   // ---------- 网络 3 ----------
   // 标题：******************************         Total Cmd . Start      ********************************
   // 含义：将 ((#Cmd.Man.StartTest OR #Step.Main.Start) AND #ManMode) AND NOT (#Step.Main.End) 赋给 #Step.Main.Start
   #Step.Main.Start := ((#Cmd.Man.StartTest OR #Step.Main.Start) AND #ManMode) AND NOT (#Step.Main.End);
   // 含义：将 ((#Cmd.Man.StartTest OR #Step.Main.Start) AND #ManMode) AND NOT (#Step.Main.End) 赋给 #Status.Busy
   #Status.Busy := ((#Cmd.Man.StartTest OR #Step.Main.Start) AND #ManMode) AND NOT (#Step.Main.End);
   // 含义：条件 NOT (((#Cmd.Man.StartTest OR #Step.Main.Start) AND #ManMode) AND NOT (#Step.Main.End)) 成立时，将 FALSE 传送到 #Status.TaskDone
   IF NOT (((#Cmd.Man.StartTest OR #Step.Main.Start) AND #ManMode) AND NOT (#Step.Main.End)) THEN
       #Status.TaskDone := FALSE;
   END_IF;
   // 含义：条件 NOT (((#Cmd.Man.StartTest OR #Step.Main.Start) AND #ManMode) AND NOT (#Step.Main.End)) 成立时，将 FALSE 传送到 #Step.Main.ErrEnd
   IF NOT (((#Cmd.Man.StartTest OR #Step.Main.Start) AND #ManMode) AND NOT (#Step.Main.End)) THEN
       #Step.Main.ErrEnd := FALSE;
   END_IF;
   // 含义：条件 NOT (((#Cmd.Man.StartTest OR #Step.Main.Start) AND #ManMode) AND NOT (#Step.Main.End)) 成立时，将 0 传送到 #Step.RandomStepNO
   IF NOT (((#Cmd.Man.StartTest OR #Step.Main.Start) AND #ManMode) AND NOT (#Step.Main.End)) THEN
       #Step.RandomStepNO := 0;
   END_IF;

   // ---------- 网络 4 ----------
   // 标题：TimeOut
   // 含义：条件 #Status.Busy AND NOT (#Step.Main.S1) 成立时，将 FALSE 传送到 #Timer_TimeOut.IN
   IF #Status.Busy AND NOT (#Step.Main.S1) THEN
       #Timer_TimeOut.IN := FALSE;
   END_IF;
   // 含义：调用定时器实例 #Timer_TimeOut
   #Timer_TimeOut(TV := #Ctrl_IN.InitParameter.TimeOutSetValue);
   // 含义：当 #Status.Busy 为 TRUE 时置位 #Timer_TimeOut.IN，否则复位（触点→线圈）
   IF #Status.Busy THEN
       #Timer_TimeOut.IN := TRUE;
   ELSE
       #Timer_TimeOut.IN := FALSE;
   END_IF;
   // 含义：条件 #Status.Busy AND #Step.Main.RandomTestCycleReStart 成立时，将 "SyS_Time" 传送到 #Aux.CycleTime_StartTime
   IF #Status.Busy AND #Step.Main.RandomTestCycleReStart THEN
       #Aux.CycleTime_StartTime := "SyS_Time";
   END_IF;
   // 含义：条件 #Status.Busy 成立时，将 ("SyS_Time" - #Aux.CycleTime_StartTime) 传送到 #Ctrl_Out.LastCylceTime
   IF #Status.Busy THEN
       #Ctrl_Out.LastCylceTime := ("SyS_Time" - #Aux.CycleTime_StartTime);
   END_IF;

   // ---------- 网络 5 ----------
   // 标题：Init
   // 含义：条件 #Step.Main.Start AND NOT (#Step.Main.S1) 成立时，将 TRUE 传送到 #Step.Main.RandomTestCycleReStart
   IF #Step.Main.Start AND NOT (#Step.Main.S1) THEN
       #Step.Main.RandomTestCycleReStart := TRUE;
   END_IF;
   // 含义：条件 #Step.Main.Start AND NOT (#Step.Main.S1) 成立时，将 #Servo_CTRL_IN.InitParameter.TimeOutSetValue 传送到 #Aux.TimeOutSetValue
   IF #Step.Main.Start AND NOT (#Step.Main.S1) THEN
       #Aux.TimeOutSetValue := #Servo_CTRL_IN.InitParameter.TimeOutSetValue;
   END_IF;
   // 含义：条件 #Step.Main.Start AND NOT (#Step.Main.S1) 成立时，将 t#15d 传送到 #Servo_CTRL_IN.InitParameter.TimeOutSetValue
   IF #Step.Main.Start AND NOT (#Step.Main.S1) THEN
       #Servo_CTRL_IN.InitParameter.TimeOutSetValue := t#15d;
   END_IF;
   // 含义：条件 #Step.Main.Start AND NOT (#Step.Main.S1) 成立时，将 0 传送到 #Ctrl_Out.AcutalCycleCounter
   IF #Step.Main.Start AND NOT (#Step.Main.S1) THEN
       #Ctrl_Out.AcutalCycleCounter := 0;
   END_IF;
   // 含义：条件 #Step.Main.Start AND NOT (#Step.Main.S1) 成立时，将 0 传送到 #Step.RandomStepNO
   IF #Step.Main.Start AND NOT (#Step.Main.S1) THEN
       #Step.RandomStepNO := 0;
   END_IF;
   // 含义：当 #Step.Main.Start 为 TRUE 时置位 #Step.Main.S1，否则复位（触点→线圈）
   IF #Step.Main.Start THEN
       #Step.Main.S1 := TRUE;
   ELSE
       #Step.Main.S1 := FALSE;
   END_IF;

   // ---------- 网络 6 ----------
   // 标题：***************************以上无需修改  ********************************
   // （空白网络）

   // ---------- 网络 7 ----------
   // 标题：乱序随机测试---随机数的生成；
   // 含义：条件 #Step.Main.RandomTestCycleReStart 成立时，将 #Step.RandomStepNO 传送到 #Ctrl_Out.LastStep
   IF #Step.Main.RandomTestCycleReStart THEN
       #Ctrl_Out.LastStep := #Step.RandomStepNO;
   END_IF;
   // 含义：条件 #Step.Main.RandomTestCycleReStart 成立时，将 (TOD_TO_DINT("SyS_Time") MOD 2) 传送到 #T_DINT
   IF #Step.Main.RandomTestCycleReStart THEN
       #T_DINT := (TOD_TO_DINT("SyS_Time") MOD 2);
   END_IF;
   // 含义：条件 #Step.Main.RandomTestCycleReStart 成立时，将 #T_DINT 传送到 #Step.RandomStepNO
   IF #Step.Main.RandomTestCycleReStart THEN
       #Step.RandomStepNO := #T_DINT;
   END_IF;
   // 含义：条件 #Step.Main.RandomTestCycleReStart 成立时，将 FALSE 传送到 #Status.TaskDone
   IF #Step.Main.RandomTestCycleReStart THEN
       #Status.TaskDone := FALSE;
   END_IF;
   // 含义：条件 #Step.Main.RandomTestCycleReStart 成立时，将 FALSE 传送到 #Status.TaskIO
   IF #Step.Main.RandomTestCycleReStart THEN
       #Status.TaskIO := FALSE;
   END_IF;

   // ---------- 网络 8 ----------
   // 标题：根据随机数进行跳转；
   // JmpList resolved

   // ---------- 网络 9 ----------
   // 标题：#Step.RandomStepNO  = 0:
   // 含义：将 ((((#Step.Main.Start AND (#Step.RandomStepNO = 0))) AND NOT (#Step.Main.RandomTestCycleReStart)) AND NOT (#Servo_Status.Busy)) OR ((((#Step.Main.Start AND (#Step.RandomStepNO = 0))) AND NOT (#Step.Main.RandomTestCycleReStart)) AND #Step.Main.S10) 赋给 #Step.Main.S10
   #Step.Main.S10 := ((((#Step.Main.Start AND (#Step.RandomStepNO = 0))) AND NOT (#Step.Main.RandomTestCycleReStart)) AND NOT (#Servo_Status.Busy)) OR ((((#Step.Main.Start AND (#Step.RandomStepNO = 0))) AND NOT (#Step.Main.RandomTestCycleReStart)) AND #Step.Main.S10);
   // 含义：条件 ((((#Step.Main.Start AND (#Step.RandomStepNO = 0))) AND NOT (#Step.Main.RandomTestCycleReStart)) AND #Step.Main.S10) AND NOT (#Step.Main.S11) 成立时，将 TRUE 传送到 #Servo_Cmd.Auto.StartTask
   IF ((((#Step.Main.Start AND (#Step.RandomStepNO = 0))) AND NOT (#Step.Main.RandomTestCycleReStart)) AND #Step.Main.S10) AND NOT (#Step.Main.S11) THEN
       #Servo_Cmd.Auto.StartTask := TRUE;
   END_IF;
   // 含义：条件 ((((#Step.Main.Start AND (#Step.RandomStepNO = 0))) AND NOT (#Step.Main.RandomTestCycleReStart)) AND #Step.Main.S10) AND NOT (#Step.Main.S11) 成立时，将 -20.0 传送到 #Servo_CTRL_IN.SetValuePosition
   IF ((((#Step.Main.Start AND (#Step.RandomStepNO = 0))) AND NOT (#Step.Main.RandomTestCycleReStart)) AND #Step.Main.S10) AND NOT (#Step.Main.S11) THEN
       #Servo_CTRL_IN.SetValuePosition := -20.0;
   END_IF;
   // 含义：将 ((((((#Step.Main.Start AND (#Step.RandomStepNO = 0))) AND NOT (#Step.Main.RandomTestCycleReStart)) AND #Step.Main.S10) AND #Servo_Status.TaskDone) AND #Servo_Status.TaskIO) OR (((((#Step.Main.Start AND (#Step.RandomStepNO = 0))) AND NOT (#Step.Main.RandomTestCycleReStart)) AND #Step.Main.S10) AND #Step.Main.S11) 赋给 #Step.Main.S11
   #Step.Main.S11 := ((((((#Step.Main.Start AND (#Step.RandomStepNO = 0))) AND NOT (#Step.Main.RandomTestCycleReStart)) AND #Step.Main.S10) AND #Servo_Status.TaskDone) AND #Servo_Status.TaskIO) OR (((((#Step.Main.Start AND (#Step.RandomStepNO = 0))) AND NOT (#Step.Main.RandomTestCycleReStart)) AND #Step.Main.S10) AND #Step.Main.S11);
   // 含义：条件 ((((((#Step.Main.Start AND (#Step.RandomStepNO = 0))) AND NOT (#Step.Main.RandomTestCycleReStart)) AND #Step.Main.S10) AND #Servo_Status.TaskDone) AND #Servo_Status.TaskIO) OR (((((#Step.Main.Start AND (#Step.RandomStepNO = 0))) AND NOT (#Step.Main.RandomTestCycleReStart)) AND #Step.Main.S10) AND #Step.Main.S11) 成立时，将 TRUE 传送到 #Status.TaskDone
   IF ((((((#Step.Main.Start AND (#Step.RandomStepNO = 0))) AND NOT (#Step.Main.RandomTestCycleReStart)) AND #Step.Main.S10) AND #Servo_Status.TaskDone) AND #Servo_Status.TaskIO) OR (((((#Step.Main.Start AND (#Step.RandomStepNO = 0))) AND NOT (#Step.Main.RandomTestCycleReStart)) AND #Step.Main.S10) AND #Step.Main.S11) THEN
       #Status.TaskDone := TRUE;
   END_IF;
   // 含义：条件 ((((((#Step.Main.Start AND (#Step.RandomStepNO = 0))) AND NOT (#Step.Main.RandomTestCycleReStart)) AND #Step.Main.S10) AND #Servo_Status.TaskDone) AND #Servo_Status.TaskIO) OR (((((#Step.Main.Start AND (#Step.RandomStepNO = 0))) AND NOT (#Step.Main.RandomTestCycleReStart)) AND #Step.Main.S10) AND #Step.Main.S11) 成立时，将 TRUE 传送到 #Status.TaskIO
   IF ((((((#Step.Main.Start AND (#Step.RandomStepNO = 0))) AND NOT (#Step.Main.RandomTestCycleReStart)) AND #Step.Main.S10) AND #Servo_Status.TaskDone) AND #Servo_Status.TaskIO) OR (((((#Step.Main.Start AND (#Step.RandomStepNO = 0))) AND NOT (#Step.Main.RandomTestCycleReStart)) AND #Step.Main.S10) AND #Step.Main.S11) THEN
       #Status.TaskIO := TRUE;
   END_IF;
   // 含义：条件 ((((((#Step.Main.Start AND (#Step.RandomStepNO = 0))) AND NOT (#Step.Main.RandomTestCycleReStart)) AND #Step.Main.S10) AND NOT (#Step.Main.S11)) AND #Servo_Status.TaskDone) AND #ErrRst 成立时，将 TRUE 传送到 #Step.Main.ErrEnd
   IF ((((((#Step.Main.Start AND (#Step.RandomStepNO = 0))) AND NOT (#Step.Main.RandomTestCycleReStart)) AND #Step.Main.S10) AND NOT (#Step.Main.S11)) AND #Servo_Status.TaskDone) AND #ErrRst THEN
       #Step.Main.ErrEnd := TRUE;
   END_IF;
   // 含义：执行该语句
   IF #Step.Main.Start THEN
       GOTO Jump;
   END_IF;

   // ---------- 网络 10 ----------
   // 标题：#Step.RandomStepNO  = 1:
   // 含义：将 ((((#Step.RandomStepNO = 1) AND #Step.Main.Start) AND NOT (#Step.Main.RandomTestCycleReStart)) AND NOT (#Servo_Status.Busy)) OR ((((#Step.RandomStepNO = 1) AND #Step.Main.Start) AND NOT (#Step.Main.RandomTestCycleReStart)) AND #Step.Main.S10) 赋给 #Step.Main.S10
   #Step.Main.S10 := ((((#Step.RandomStepNO = 1) AND #Step.Main.Start) AND NOT (#Step.Main.RandomTestCycleReStart)) AND NOT (#Servo_Status.Busy)) OR ((((#Step.RandomStepNO = 1) AND #Step.Main.Start) AND NOT (#Step.Main.RandomTestCycleReStart)) AND #Step.Main.S10);
   // 含义：条件 ((((#Step.RandomStepNO = 1) AND #Step.Main.Start) AND NOT (#Step.Main.RandomTestCycleReStart)) AND #Step.Main.S10) AND NOT (#Step.Main.S11) 成立时，将 TRUE 传送到 #Servo_Cmd.Auto.StartTask
   IF ((((#Step.RandomStepNO = 1) AND #Step.Main.Start) AND NOT (#Step.Main.RandomTestCycleReStart)) AND #Step.Main.S10) AND NOT (#Step.Main.S11) THEN
       #Servo_Cmd.Auto.StartTask := TRUE;
   END_IF;
   // 含义：条件 ((((#Step.RandomStepNO = 1) AND #Step.Main.Start) AND NOT (#Step.Main.RandomTestCycleReStart)) AND #Step.Main.S10) AND NOT (#Step.Main.S11) 成立时，将 20.0 传送到 #Servo_CTRL_IN.SetValuePosition
   IF ((((#Step.RandomStepNO = 1) AND #Step.Main.Start) AND NOT (#Step.Main.RandomTestCycleReStart)) AND #Step.Main.S10) AND NOT (#Step.Main.S11) THEN
       #Servo_CTRL_IN.SetValuePosition := 20.0;
   END_IF;
   // 含义：将 ((((((#Step.RandomStepNO = 1) AND #Step.Main.Start) AND NOT (#Step.Main.RandomTestCycleReStart)) AND #Step.Main.S10) AND #Servo_Status.TaskDone) AND #Servo_Status.TaskIO) OR (((((#Step.RandomStepNO = 1) AND #Step.Main.Start) AND NOT (#Step.Main.RandomTestCycleReStart)) AND #Step.Main.S10) AND #Step.Main.S11) 赋给 #Step.Main.S11
   #Step.Main.S11 := ((((((#Step.RandomStepNO = 1) AND #Step.Main.Start) AND NOT (#Step.Main.RandomTestCycleReStart)) AND #Step.Main.S10) AND #Servo_Status.TaskDone) AND #Servo_Status.TaskIO) OR (((((#Step.RandomStepNO = 1) AND #Step.Main.Start) AND NOT (#Step.Main.RandomTestCycleReStart)) AND #Step.Main.S10) AND #Step.Main.S11);
   // 含义：条件 ((((((#Step.RandomStepNO = 1) AND #Step.Main.Start) AND NOT (#Step.Main.RandomTestCycleReStart)) AND #Step.Main.S10) AND #Servo_Status.TaskDone) AND #Servo_Status.TaskIO) OR (((((#Step.RandomStepNO = 1) AND #Step.Main.Start) AND NOT (#Step.Main.RandomTestCycleReStart)) AND #Step.Main.S10) AND #Step.Main.S11) 成立时，将 TRUE 传送到 #Status.TaskDone
   IF ((((((#Step.RandomStepNO = 1) AND #Step.Main.Start) AND NOT (#Step.Main.RandomTestCycleReStart)) AND #Step.Main.S10) AND #Servo_Status.TaskDone) AND #Servo_Status.TaskIO) OR (((((#Step.RandomStepNO = 1) AND #Step.Main.Start) AND NOT (#Step.Main.RandomTestCycleReStart)) AND #Step.Main.S10) AND #Step.Main.S11) THEN
       #Status.TaskDone := TRUE;
   END_IF;
   // 含义：条件 ((((((#Step.RandomStepNO = 1) AND #Step.Main.Start) AND NOT (#Step.Main.RandomTestCycleReStart)) AND #Step.Main.S10) AND #Servo_Status.TaskDone) AND #Servo_Status.TaskIO) OR (((((#Step.RandomStepNO = 1) AND #Step.Main.Start) AND NOT (#Step.Main.RandomTestCycleReStart)) AND #Step.Main.S10) AND #Step.Main.S11) 成立时，将 TRUE 传送到 #Status.TaskIO
   IF ((((((#Step.RandomStepNO = 1) AND #Step.Main.Start) AND NOT (#Step.Main.RandomTestCycleReStart)) AND #Step.Main.S10) AND #Servo_Status.TaskDone) AND #Servo_Status.TaskIO) OR (((((#Step.RandomStepNO = 1) AND #Step.Main.Start) AND NOT (#Step.Main.RandomTestCycleReStart)) AND #Step.Main.S10) AND #Step.Main.S11) THEN
       #Status.TaskIO := TRUE;
   END_IF;
   // 含义：条件 ((((((#Step.RandomStepNO = 1) AND #Step.Main.Start) AND NOT (#Step.Main.RandomTestCycleReStart)) AND #Step.Main.S10) AND NOT (#Step.Main.S11)) AND #Servo_Status.TaskDone) AND #ErrRst 成立时，将 TRUE 传送到 #Step.Main.ErrEnd
   IF ((((((#Step.RandomStepNO = 1) AND #Step.Main.Start) AND NOT (#Step.Main.RandomTestCycleReStart)) AND #Step.Main.S10) AND NOT (#Step.Main.S11)) AND #Servo_Status.TaskDone) AND #ErrRst THEN
       #Step.Main.ErrEnd := TRUE;
   END_IF;
   // 含义：执行该语句
   IF (#Step.RandomStepNO = 1) AND #Step.Main.Start THEN
       GOTO Jump;
   END_IF;

   // ---------- 网络 11 ----------
   // 标题：#Step.RandomStepNO  = 2:
   // 含义：将 ((((#Step.Main.Start AND (#Step.RandomStepNO = 2))) AND NOT (#Step.Main.RandomTestCycleReStart)) AND NOT (#Servo_Status.Busy)) OR ((((#Step.Main.Start AND (#Step.RandomStepNO = 2))) AND NOT (#Step.Main.RandomTestCycleReStart)) AND #Step.Main.S10) 赋给 #Step.Main.S10
   #Step.Main.S10 := ((((#Step.Main.Start AND (#Step.RandomStepNO = 2))) AND NOT (#Step.Main.RandomTestCycleReStart)) AND NOT (#Servo_Status.Busy)) OR ((((#Step.Main.Start AND (#Step.RandomStepNO = 2))) AND NOT (#Step.Main.RandomTestCycleReStart)) AND #Step.Main.S10);
   // 含义：条件 ((((#Step.Main.Start AND (#Step.RandomStepNO = 2))) AND NOT (#Step.Main.RandomTestCycleReStart)) AND #Step.Main.S10) AND NOT (#Step.Main.S11) 成立时，将 TRUE 传送到 #Servo_Cmd.Auto.StartTask_TLM
   IF ((((#Step.Main.Start AND (#Step.RandomStepNO = 2))) AND NOT (#Step.Main.RandomTestCycleReStart)) AND #Step.Main.S10) AND NOT (#Step.Main.S11) THEN
       #Servo_Cmd.Auto.StartTask_TLM := TRUE;
   END_IF;
   // 含义：条件 ((((#Step.Main.Start AND (#Step.RandomStepNO = 2))) AND NOT (#Step.Main.RandomTestCycleReStart)) AND #Step.Main.S10) AND NOT (#Step.Main.S11) 成立时，将 10.0 传送到 #Servo_CTRL_IN.SetValuePosition
   IF ((((#Step.Main.Start AND (#Step.RandomStepNO = 2))) AND NOT (#Step.Main.RandomTestCycleReStart)) AND #Step.Main.S10) AND NOT (#Step.Main.S11) THEN
       #Servo_CTRL_IN.SetValuePosition := 10.0;
   END_IF;
   // 含义：将 ((((((#Step.Main.Start AND (#Step.RandomStepNO = 2))) AND NOT (#Step.Main.RandomTestCycleReStart)) AND #Step.Main.S10) AND #Servo_Status.TaskDone) AND #Servo_Status.TaskIO) OR (((((#Step.Main.Start AND (#Step.RandomStepNO = 2))) AND NOT (#Step.Main.RandomTestCycleReStart)) AND #Step.Main.S10) AND #Step.Main.S11) 赋给 #Step.Main.S11
   #Step.Main.S11 := ((((((#Step.Main.Start AND (#Step.RandomStepNO = 2))) AND NOT (#Step.Main.RandomTestCycleReStart)) AND #Step.Main.S10) AND #Servo_Status.TaskDone) AND #Servo_Status.TaskIO) OR (((((#Step.Main.Start AND (#Step.RandomStepNO = 2))) AND NOT (#Step.Main.RandomTestCycleReStart)) AND #Step.Main.S10) AND #Step.Main.S11);
   // 含义：条件 ((((((#Step.Main.Start AND (#Step.RandomStepNO = 2))) AND NOT (#Step.Main.RandomTestCycleReStart)) AND #Step.Main.S10) AND #Servo_Status.TaskDone) AND #Servo_Status.TaskIO) OR (((((#Step.Main.Start AND (#Step.RandomStepNO = 2))) AND NOT (#Step.Main.RandomTestCycleReStart)) AND #Step.Main.S10) AND #Step.Main.S11) 成立时，将 TRUE 传送到 #Status.TaskDone
   IF ((((((#Step.Main.Start AND (#Step.RandomStepNO = 2))) AND NOT (#Step.Main.RandomTestCycleReStart)) AND #Step.Main.S10) AND #Servo_Status.TaskDone) AND #Servo_Status.TaskIO) OR (((((#Step.Main.Start AND (#Step.RandomStepNO = 2))) AND NOT (#Step.Main.RandomTestCycleReStart)) AND #Step.Main.S10) AND #Step.Main.S11) THEN
       #Status.TaskDone := TRUE;
   END_IF;
   // 含义：条件 ((((((#Step.Main.Start AND (#Step.RandomStepNO = 2))) AND NOT (#Step.Main.RandomTestCycleReStart)) AND #Step.Main.S10) AND #Servo_Status.TaskDone) AND #Servo_Status.TaskIO) OR (((((#Step.Main.Start AND (#Step.RandomStepNO = 2))) AND NOT (#Step.Main.RandomTestCycleReStart)) AND #Step.Main.S10) AND #Step.Main.S11) 成立时，将 TRUE 传送到 #Status.TaskIO
   IF ((((((#Step.Main.Start AND (#Step.RandomStepNO = 2))) AND NOT (#Step.Main.RandomTestCycleReStart)) AND #Step.Main.S10) AND #Servo_Status.TaskDone) AND #Servo_Status.TaskIO) OR (((((#Step.Main.Start AND (#Step.RandomStepNO = 2))) AND NOT (#Step.Main.RandomTestCycleReStart)) AND #Step.Main.S10) AND #Step.Main.S11) THEN
       #Status.TaskIO := TRUE;
   END_IF;
   // 含义：条件 ((((((#Step.Main.Start AND (#Step.RandomStepNO = 2))) AND NOT (#Step.Main.RandomTestCycleReStart)) AND #Step.Main.S10) AND NOT (#Step.Main.S11)) AND #Servo_Status.TaskDone) AND #ErrRst 成立时，将 TRUE 传送到 #Step.Main.ErrEnd
   IF ((((((#Step.Main.Start AND (#Step.RandomStepNO = 2))) AND NOT (#Step.Main.RandomTestCycleReStart)) AND #Step.Main.S10) AND NOT (#Step.Main.S11)) AND #Servo_Status.TaskDone) AND #ErrRst THEN
       #Step.Main.ErrEnd := TRUE;
   END_IF;
   // 含义：执行该语句
   IF #Step.Main.Start THEN
       GOTO Jump;
   END_IF;

   // ---------- 网络 12 ----------
   // 标题：#Step.RandomStepNO  = 3:
   // 含义：将 ((((#Step.Main.Start AND (#Step.RandomStepNO = 3))) AND NOT (#Step.Main.RandomTestCycleReStart)) AND NOT (#Servo_Status.Busy)) OR ((((#Step.Main.Start AND (#Step.RandomStepNO = 3))) AND NOT (#Step.Main.RandomTestCycleReStart)) AND #Step.Main.S10) 赋给 #Step.Main.S10
   #Step.Main.S10 := ((((#Step.Main.Start AND (#Step.RandomStepNO = 3))) AND NOT (#Step.Main.RandomTestCycleReStart)) AND NOT (#Servo_Status.Busy)) OR ((((#Step.Main.Start AND (#Step.RandomStepNO = 3))) AND NOT (#Step.Main.RandomTestCycleReStart)) AND #Step.Main.S10);
   // 含义：条件 ((((#Step.Main.Start AND (#Step.RandomStepNO = 3))) AND NOT (#Step.Main.RandomTestCycleReStart)) AND #Step.Main.S10) AND NOT (#Step.Main.S11) 成立时，将 TRUE 传送到 #Servo_Cmd.Auto.SetTLM
   IF ((((#Step.Main.Start AND (#Step.RandomStepNO = 3))) AND NOT (#Step.Main.RandomTestCycleReStart)) AND #Step.Main.S10) AND NOT (#Step.Main.S11) THEN
       #Servo_Cmd.Auto.SetTLM := TRUE;
   END_IF;
   // 含义：将 ((((((#Step.Main.Start AND (#Step.RandomStepNO = 3))) AND NOT (#Step.Main.RandomTestCycleReStart)) AND #Step.Main.S10) AND #Servo_Status.TaskDone) AND #Servo_Status.TaskIO) OR (((((#Step.Main.Start AND (#Step.RandomStepNO = 3))) AND NOT (#Step.Main.RandomTestCycleReStart)) AND #Step.Main.S10) AND #Step.Main.S11) 赋给 #Step.Main.S11
   #Step.Main.S11 := ((((((#Step.Main.Start AND (#Step.RandomStepNO = 3))) AND NOT (#Step.Main.RandomTestCycleReStart)) AND #Step.Main.S10) AND #Servo_Status.TaskDone) AND #Servo_Status.TaskIO) OR (((((#Step.Main.Start AND (#Step.RandomStepNO = 3))) AND NOT (#Step.Main.RandomTestCycleReStart)) AND #Step.Main.S10) AND #Step.Main.S11);
   // 含义：条件 ((((((#Step.Main.Start AND (#Step.RandomStepNO = 3))) AND NOT (#Step.Main.RandomTestCycleReStart)) AND #Step.Main.S10) AND #Servo_Status.TaskDone) AND #Servo_Status.TaskIO) OR (((((#Step.Main.Start AND (#Step.RandomStepNO = 3))) AND NOT (#Step.Main.RandomTestCycleReStart)) AND #Step.Main.S10) AND #Step.Main.S11) 成立时，将 TRUE 传送到 #Status.TaskDone
   IF ((((((#Step.Main.Start AND (#Step.RandomStepNO = 3))) AND NOT (#Step.Main.RandomTestCycleReStart)) AND #Step.Main.S10) AND #Servo_Status.TaskDone) AND #Servo_Status.TaskIO) OR (((((#Step.Main.Start AND (#Step.RandomStepNO = 3))) AND NOT (#Step.Main.RandomTestCycleReStart)) AND #Step.Main.S10) AND #Step.Main.S11) THEN
       #Status.TaskDone := TRUE;
   END_IF;
   // 含义：条件 ((((((#Step.Main.Start AND (#Step.RandomStepNO = 3))) AND NOT (#Step.Main.RandomTestCycleReStart)) AND #Step.Main.S10) AND #Servo_Status.TaskDone) AND #Servo_Status.TaskIO) OR (((((#Step.Main.Start AND (#Step.RandomStepNO = 3))) AND NOT (#Step.Main.RandomTestCycleReStart)) AND #Step.Main.S10) AND #Step.Main.S11) 成立时，将 TRUE 传送到 #Status.TaskIO
   IF ((((((#Step.Main.Start AND (#Step.RandomStepNO = 3))) AND NOT (#Step.Main.RandomTestCycleReStart)) AND #Step.Main.S10) AND #Servo_Status.TaskDone) AND #Servo_Status.TaskIO) OR (((((#Step.Main.Start AND (#Step.RandomStepNO = 3))) AND NOT (#Step.Main.RandomTestCycleReStart)) AND #Step.Main.S10) AND #Step.Main.S11) THEN
       #Status.TaskIO := TRUE;
   END_IF;
   // 含义：条件 ((((((#Step.Main.Start AND (#Step.RandomStepNO = 3))) AND NOT (#Step.Main.RandomTestCycleReStart)) AND #Step.Main.S10) AND NOT (#Step.Main.S11)) AND #Servo_Status.TaskDone) AND #ErrRst 成立时，将 TRUE 传送到 #Step.Main.ErrEnd
   IF ((((((#Step.Main.Start AND (#Step.RandomStepNO = 3))) AND NOT (#Step.Main.RandomTestCycleReStart)) AND #Step.Main.S10) AND NOT (#Step.Main.S11)) AND #Servo_Status.TaskDone) AND #ErrRst THEN
       #Step.Main.ErrEnd := TRUE;
   END_IF;
   // 含义：执行该语句
   IF #Step.Main.Start THEN
       GOTO Jump;
   END_IF;

   // ---------- 网络 13 ----------
   // 标题：#Step.RandomStepNO  = 4:
   // 含义：将 ((((#Step.Main.Start AND (#Step.RandomStepNO = 4))) AND NOT (#Step.Main.RandomTestCycleReStart)) AND NOT (#Servo_Status.Busy)) OR ((((#Step.Main.Start AND (#Step.RandomStepNO = 4))) AND NOT (#Step.Main.RandomTestCycleReStart)) AND #Step.Main.S10) 赋给 #Step.Main.S10
   #Step.Main.S10 := ((((#Step.Main.Start AND (#Step.RandomStepNO = 4))) AND NOT (#Step.Main.RandomTestCycleReStart)) AND NOT (#Servo_Status.Busy)) OR ((((#Step.Main.Start AND (#Step.RandomStepNO = 4))) AND NOT (#Step.Main.RandomTestCycleReStart)) AND #Step.Main.S10);
   // 含义：条件 ((((#Step.Main.Start AND (#Step.RandomStepNO = 4))) AND NOT (#Step.Main.RandomTestCycleReStart)) AND #Step.Main.S10) AND NOT (#Step.Main.S11) 成立时，将 TRUE 传送到 #Servo_Cmd.Auto.JogPos
   IF ((((#Step.Main.Start AND (#Step.RandomStepNO = 4))) AND NOT (#Step.Main.RandomTestCycleReStart)) AND #Step.Main.S10) AND NOT (#Step.Main.S11) THEN
       #Servo_Cmd.Auto.JogPos := TRUE;
   END_IF;
   // 含义：将 ((((((#Step.Main.Start AND (#Step.RandomStepNO = 4))) AND NOT (#Step.Main.RandomTestCycleReStart)) AND #Step.Main.S10) AND (#Servo_CTRL_OUT.ActualPosition >= 10.0))) OR (((((#Step.Main.Start AND (#Step.RandomStepNO = 4))) AND NOT (#Step.Main.RandomTestCycleReStart)) AND #Step.Main.S10) AND #Step.Main.S11) 赋给 #Step.Main.S11
   #Step.Main.S11 := ((((((#Step.Main.Start AND (#Step.RandomStepNO = 4))) AND NOT (#Step.Main.RandomTestCycleReStart)) AND #Step.Main.S10) AND (#Servo_CTRL_OUT.ActualPosition >= 10.0))) OR (((((#Step.Main.Start AND (#Step.RandomStepNO = 4))) AND NOT (#Step.Main.RandomTestCycleReStart)) AND #Step.Main.S10) AND #Step.Main.S11);
   // 含义：条件 ((((((#Step.Main.Start AND (#Step.RandomStepNO = 4))) AND NOT (#Step.Main.RandomTestCycleReStart)) AND #Step.Main.S10) AND (#Servo_CTRL_OUT.ActualPosition >= 10.0))) OR (((((#Step.Main.Start AND (#Step.RandomStepNO = 4))) AND NOT (#Step.Main.RandomTestCycleReStart)) AND #Step.Main.S10) AND #Step.Main.S11) 成立时，将 TRUE 传送到 #Status.TaskDone
   IF ((((((#Step.Main.Start AND (#Step.RandomStepNO = 4))) AND NOT (#Step.Main.RandomTestCycleReStart)) AND #Step.Main.S10) AND (#Servo_CTRL_OUT.ActualPosition >= 10.0))) OR (((((#Step.Main.Start AND (#Step.RandomStepNO = 4))) AND NOT (#Step.Main.RandomTestCycleReStart)) AND #Step.Main.S10) AND #Step.Main.S11) THEN
       #Status.TaskDone := TRUE;
   END_IF;
   // 含义：条件 ((((((#Step.Main.Start AND (#Step.RandomStepNO = 4))) AND NOT (#Step.Main.RandomTestCycleReStart)) AND #Step.Main.S10) AND (#Servo_CTRL_OUT.ActualPosition >= 10.0))) OR (((((#Step.Main.Start AND (#Step.RandomStepNO = 4))) AND NOT (#Step.Main.RandomTestCycleReStart)) AND #Step.Main.S10) AND #Step.Main.S11) 成立时，将 TRUE 传送到 #Status.TaskIO
   IF ((((((#Step.Main.Start AND (#Step.RandomStepNO = 4))) AND NOT (#Step.Main.RandomTestCycleReStart)) AND #Step.Main.S10) AND (#Servo_CTRL_OUT.ActualPosition >= 10.0))) OR (((((#Step.Main.Start AND (#Step.RandomStepNO = 4))) AND NOT (#Step.Main.RandomTestCycleReStart)) AND #Step.Main.S10) AND #Step.Main.S11) THEN
       #Status.TaskIO := TRUE;
   END_IF;
   // 含义：条件 ((((((#Step.Main.Start AND (#Step.RandomStepNO = 4))) AND NOT (#Step.Main.RandomTestCycleReStart)) AND #Step.Main.S10) AND NOT (#Step.Main.S11)) AND #Servo_Status.TaskDone) AND #ErrRst 成立时，将 TRUE 传送到 #Step.Main.ErrEnd
   IF ((((((#Step.Main.Start AND (#Step.RandomStepNO = 4))) AND NOT (#Step.Main.RandomTestCycleReStart)) AND #Step.Main.S10) AND NOT (#Step.Main.S11)) AND #Servo_Status.TaskDone) AND #ErrRst THEN
       #Step.Main.ErrEnd := TRUE;
   END_IF;
   // 含义：执行该语句
   IF #Step.Main.Start THEN
       GOTO Jump;
   END_IF;

   // ---------- 网络 14 ----------
   // 标题：#Step.RandomStepNO  = 4:
   // 含义：将 ((((#Step.Main.Start AND (#Step.RandomStepNO = 5))) AND NOT (#Step.Main.RandomTestCycleReStart)) AND NOT (#Servo_Status.Busy)) OR ((((#Step.Main.Start AND (#Step.RandomStepNO = 5))) AND NOT (#Step.Main.RandomTestCycleReStart)) AND #Step.Main.S10) 赋给 #Step.Main.S10
   #Step.Main.S10 := ((((#Step.Main.Start AND (#Step.RandomStepNO = 5))) AND NOT (#Step.Main.RandomTestCycleReStart)) AND NOT (#Servo_Status.Busy)) OR ((((#Step.Main.Start AND (#Step.RandomStepNO = 5))) AND NOT (#Step.Main.RandomTestCycleReStart)) AND #Step.Main.S10);
   // 含义：条件 ((((#Step.Main.Start AND (#Step.RandomStepNO = 5))) AND NOT (#Step.Main.RandomTestCycleReStart)) AND #Step.Main.S10) AND NOT (#Step.Main.S11) 成立时，将 TRUE 传送到 #Servo_Cmd.Auto.TorqueCtrl_FixedStop
   IF ((((#Step.Main.Start AND (#Step.RandomStepNO = 5))) AND NOT (#Step.Main.RandomTestCycleReStart)) AND #Step.Main.S10) AND NOT (#Step.Main.S11) THEN
       #Servo_Cmd.Auto.TorqueCtrl_FixedStop := TRUE;
   END_IF;
   // 含义：条件 ((((#Step.Main.Start AND (#Step.RandomStepNO = 5))) AND NOT (#Step.Main.RandomTestCycleReStart)) AND #Step.Main.S10) AND NOT (#Step.Main.S11) 成立时，将 50.0 传送到 #Servo_CTRL_IN.SetValuePosition
   IF ((((#Step.Main.Start AND (#Step.RandomStepNO = 5))) AND NOT (#Step.Main.RandomTestCycleReStart)) AND #Step.Main.S10) AND NOT (#Step.Main.S11) THEN
       #Servo_CTRL_IN.SetValuePosition := 50.0;
   END_IF;
   // 含义：将 ((((((#Step.Main.Start AND (#Step.RandomStepNO = 5))) AND NOT (#Step.Main.RandomTestCycleReStart)) AND #Step.Main.S10) AND #Servo_Status.TaskDone) AND #Servo_Status.TaskNIO) OR ((((((#Step.Main.Start AND (#Step.RandomStepNO = 5))) AND NOT (#Step.Main.RandomTestCycleReStart)) AND #Step.Main.S10) AND #Servo_Status.TaskDone) AND #Servo_Status.TaskIO) OR (((((#Step.Main.Start AND (#Step.RandomStepNO = 5))) AND NOT (#Step.Main.RandomTestCycleReStart)) AND #Step.Main.S10) AND #Step.Main.S11) 赋给 #Step.Main.S11
   #Step.Main.S11 := ((((((#Step.Main.Start AND (#Step.RandomStepNO = 5))) AND NOT (#Step.Main.RandomTestCycleReStart)) AND #Step.Main.S10) AND #Servo_Status.TaskDone) AND #Servo_Status.TaskNIO) OR ((((((#Step.Main.Start AND (#Step.RandomStepNO = 5))) AND NOT (#Step.Main.RandomTestCycleReStart)) AND #Step.Main.S10) AND #Servo_Status.TaskDone) AND #Servo_Status.TaskIO) OR (((((#Step.Main.Start AND (#Step.RandomStepNO = 5))) AND NOT (#Step.Main.RandomTestCycleReStart)) AND #Step.Main.S10) AND #Step.Main.S11);
   // 含义：条件 ((((#Step.Main.Start AND (#Step.RandomStepNO = 5))) AND NOT (#Step.Main.RandomTestCycleReStart)) AND #Step.Main.S11) AND NOT (#Step.Main.S12) 成立时，将 TRUE 传送到 "ErrRst_M"
   IF ((((#Step.Main.Start AND (#Step.RandomStepNO = 5))) AND NOT (#Step.Main.RandomTestCycleReStart)) AND #Step.Main.S11) AND NOT (#Step.Main.S12) THEN
       "ErrRst_M" := TRUE;
   END_IF;
   // 含义：条件 (((((#Step.Main.Start AND (#Step.RandomStepNO = 5))) AND NOT (#Step.Main.RandomTestCycleReStart)) AND #Step.Main.S11) AND NOT (#Servo_Status.TaskDone)) AND #Servo_Status.OkToStart 成立时，将 TRUE 传送到 #Status.TaskDone
   IF (((((#Step.Main.Start AND (#Step.RandomStepNO = 5))) AND NOT (#Step.Main.RandomTestCycleReStart)) AND #Step.Main.S11) AND NOT (#Servo_Status.TaskDone)) AND #Servo_Status.OkToStart THEN
       #Status.TaskDone := TRUE;
   END_IF;
   // 含义：条件 (((((#Step.Main.Start AND (#Step.RandomStepNO = 5))) AND NOT (#Step.Main.RandomTestCycleReStart)) AND #Step.Main.S11) AND NOT (#Servo_Status.TaskDone)) AND #Servo_Status.OkToStart 成立时，将 TRUE 传送到 #Status.TaskIO
   IF (((((#Step.Main.Start AND (#Step.RandomStepNO = 5))) AND NOT (#Step.Main.RandomTestCycleReStart)) AND #Step.Main.S11) AND NOT (#Servo_Status.TaskDone)) AND #Servo_Status.OkToStart THEN
       #Status.TaskIO := TRUE;
   END_IF;
   // 含义：将 (((((#Step.Main.Start AND (#Step.RandomStepNO = 5))) AND NOT (#Step.Main.RandomTestCycleReStart)) AND #Step.Main.S11) AND NOT (#Servo_Status.TaskDone)) AND #Servo_Status.OkToStart 赋给 #Step.Main.S12
   #Step.Main.S12 := (((((#Step.Main.Start AND (#Step.RandomStepNO = 5))) AND NOT (#Step.Main.RandomTestCycleReStart)) AND #Step.Main.S11) AND NOT (#Servo_Status.TaskDone)) AND #Servo_Status.OkToStart;
   // 含义：执行该语句
   IF #Step.Main.Start THEN
       GOTO Jump;
   END_IF;

   // ---------- 网络 15 ----------
   // 标题：*******************以下无需修改******************************************
   // （空白网络）

   // ---------- 网络 16 ----------
   // 标题：***************************************无条件复位***********
   // 含义：将 FALSE 赋给 #Step.Main.RandomTestCycleReStart
   Jump:
   ;

   #Step.Main.RandomTestCycleReStart := FALSE;

   // ---------- 网络 17 ----------
   // 标题：判断测试是否结束
   // 含义：条件 (#Status.TaskDone AND #Status.TaskIO) AND NOT (#Step.Main.S50) 成立时，将 (#Ctrl_Out.AcutalCycleCounter + 1) 传送到 #Ctrl_Out.AcutalCycleCounter
   IF (#Status.TaskDone AND #Status.TaskIO) AND NOT (#Step.Main.S50) THEN
       #Ctrl_Out.AcutalCycleCounter := (#Ctrl_Out.AcutalCycleCounter + 1);
   END_IF;
   // 含义：将 (((#Status.TaskDone AND #Status.TaskIO) AND (#Ctrl_Out.AcutalCycleCounter >= #Ctrl_IN.TestCycleCounter))) OR ((#Status.TaskDone AND #Status.TaskIO) AND NOT (#Cmd.Man.StartTest)) OR ((#Status.TaskDone AND #Status.TaskIO) AND #Step.Main.S50) 赋给 #Step.Main.S50
   #Step.Main.S50 := (((#Status.TaskDone AND #Status.TaskIO) AND (#Ctrl_Out.AcutalCycleCounter >= #Ctrl_IN.TestCycleCounter))) OR ((#Status.TaskDone AND #Status.TaskIO) AND NOT (#Cmd.Man.StartTest)) OR ((#Status.TaskDone AND #Status.TaskIO) AND #Step.Main.S50);
   // 含义：条件 (#Status.TaskDone AND #Status.TaskIO) AND NOT (#Step.Main.S50) 成立时，将 TRUE 传送到 #Step.Main.RandomTestCycleReStart
   IF (#Status.TaskDone AND #Status.TaskIO) AND NOT (#Step.Main.S50) THEN
       #Step.Main.RandomTestCycleReStart := TRUE;
   END_IF;

   // ---------- 网络 18 ----------
   // 标题：Wait Cmd.Off
   // 含义：当 #Step.Main.S50 为 TRUE 时置位 #Step.Main.End，否则复位（触点→线圈）
   IF #Step.Main.S50 THEN
       #Step.Main.End := TRUE;
   ELSE
       #Step.Main.End := FALSE;
   END_IF;
   // 含义：条件 #Step.Main.S50 成立时，将 0 传送到 #TP_Cmd
   IF #Step.Main.S50 THEN
       #TP_Cmd := 0;
   END_IF;

   // ---------- 网络 19 ----------
   // 标题：恢复默认的超时时间；
   // 含义：将 (#Step.Main.S1 OR #Step.Main.DTResetS1) AND NOT (#Step.Main.DTResetS2) 赋给 #Step.Main.DTResetS1
   #Step.Main.DTResetS1 := (#Step.Main.S1 OR #Step.Main.DTResetS1) AND NOT (#Step.Main.DTResetS2);
   // 含义：将 (#Step.Main.DTResetS1 AND NOT (#Step.Main.Start)) OR (#Step.Main.DTResetS1 AND #Step.Main.DTResetS2) 赋给 #Step.Main.DTResetS2
   #Step.Main.DTResetS2 := (#Step.Main.DTResetS1 AND NOT (#Step.Main.Start)) OR (#Step.Main.DTResetS1 AND #Step.Main.DTResetS2);
   // 含义：条件 (#Step.Main.DTResetS1 AND NOT (#Step.Main.Start)) OR (#Step.Main.DTResetS1 AND #Step.Main.DTResetS2) 成立时，将 #Aux.TimeOutSetValue 传送到 #Servo_CTRL_IN.InitParameter.TimeOutSetValue
   IF (#Step.Main.DTResetS1 AND NOT (#Step.Main.Start)) OR (#Step.Main.DTResetS1 AND #Step.Main.DTResetS2) THEN
       #Servo_CTRL_IN.InitParameter.TimeOutSetValue := #Aux.TimeOutSetValue;
   END_IF;
END_FUNCTION_BLOCK

FUNCTION_BLOCK "FB5715_Kuka_General"   // FB5715, SCL
{ S7_Optimized_Access := 'TRUE' }
// ============================================================
//  Block: FB5715_Kuka_General
//  ============================================================
//  编号：FB5715
//  原始语言：SCL（规则翻译为 SCL）
//  含义：2019.09.25
//  1.用于Yamaha-TS系列PN接口的单轴伺服
   VAR_INPUT
      ManMode : Bool;   // 输入参数
      AllMode : Bool;   // 输入参数
      EMMode : Bool;   // 输入参数
      ErrRst : Bool;   // 输入参数
      RobotEnble : Bool;   // 使能信号
      PromptStruct : Struct   // 输入参数
         Info : Struct   // 输入参数
            bit0 : Bool;   // 输入参数
            bit1 : Bool;   // 输入参数
            bit2 : Bool;   // 输入参数
            bit3 : Bool;   // 输入参数
            bit4 : Bool;   // 输入参数
            bit5 : Bool;   // 输入参数
            bit6 : Bool;   // 输入参数
            bit7 : Bool;   // 输入参数
            bit8 : Bool;   // 输入参数
            bit9 : Bool;   // 输入参数
            bit10 : Bool;   // 输入参数
            bit11 : Bool;   // 输入参数
            bit12 : Bool;   // 输入参数
            bit13 : Bool;   // 输入参数
            bit14 : Bool;   // 输入参数
            bit15 : Bool;   // 输入参数
            bit16 : Bool;   // 输入参数
            bit17 : Bool;   // 输入参数
            bit18 : Bool;   // 输入参数
            bit19 : Bool;   // 输入参数
            bit20 : Bool;   // 输入参数
            bit21 : Bool;   // 输入参数
            bit22 : Bool;   // 输入参数
            bit23 : Bool;   // 输入参数
            bit24 : Bool;   // 输入参数
            bit25 : Bool;   // 输入参数
            bit26 : Bool;   // 输入参数
            bit27 : Bool;   // 输入参数
            bit28 : Bool;   // 输入参数
            bit29 : Bool;   // 输入参数
            bit30 : Bool;   // 输入参数
            bit31 : Bool;   // 输入参数
         END_STRUCT;
         Err : Struct   // 输入参数
            bit0 : Bool;   // 输入参数
            bit1 : Bool;   // 输入参数
            bit2 : Bool;   // 输入参数
            bit3 : Bool;   // 输入参数
            bit4 : Bool;   // 输入参数
            bit5 : Bool;   // 输入参数
            bit6 : Bool;   // 输入参数
            bit7 : Bool;   // 输入参数
            bit8 : Bool;   // 输入参数
            bit9 : Bool;   // 输入参数
            bit10 : Bool;   // 输入参数
            bit11 : Bool;   // 输入参数
            bit12 : Bool;   // 输入参数
            bit13 : Bool;   // 输入参数
            bit14 : Bool;   // 输入参数
            bit15 : Bool;   // 输入参数
            bit16 : Bool;   // 输入参数
            bit17 : Bool;   // 输入参数
            bit18 : Bool;   // 输入参数
            bit19 : Bool;   // 输入参数
            bit20 : Bool;   // 输入参数
            bit21 : Bool;   // 输入参数
            bit22 : Bool;   // 输入参数
            bit23 : Bool;   // 输入参数
            bit24 : Bool;   // 输入参数
            bit25 : Bool;   // 输入参数
            bit26 : Bool;   // 输入参数
            bit27 : Bool;   // 输入参数
            bit28 : Bool;   // 输入参数
            bit29 : Bool;   // 输入参数
            bit30 : Bool;   // 输入参数
            bit31 : Bool;   // 输入参数
         END_STRUCT;
      END_STRUCT;
      IN : Bool;   // 输入参数
      TV : Time;   // 输入参数
   END_VAR
   VAR_OUTPUT
      PromptValue : Int;   // 输出参数
      Q : Bool;   // 输出参数
   END_VAR
   VAR
      TP_Cmd : Word;   // 用于触摸屏操作
      TP_Status : Word;   // 静态变量
      Cmd : Struct   // 静态变量
         Auto : Struct   // 静态变量
            ProgStart : Bool;   // 静态变量
            GoHome : Bool;   // 静态变量
            Stop : Bool;   // 静态变量
         END_STRUCT;
      END_STRUCT;
      AtCmd : Struct   // 静态变量
         Auto : Word;   // 静态变量
      END_STRUCT;
      CTRL_IN : Struct   // in控制用数据接口：8
         ProgNo : Byte;   // 程序号
         RobotSpeed : Byte;   // 机器人速度
         InitParameter : Struct   // 静态变量
            HW_Addr : Hw_Io := 999;   // IO地址或者硬件标识符
            TimeOutSetValue : Time := T#16M_40S;   // 默认--15S内，命令必须能正常结束；
            Td : Time := T#5MS;   // 默认参数，5ms，指令识别延时
            sp : Array[0..3] of Real;   // 静态变量
         END_STRUCT;
      END_STRUCT;
      CTRL_OUT : Struct   // out控制用数据接口：60
         ProgNo : Byte;   // 程序号
         AppInfNo : Byte;   // 操作提示
         ErrorCode : Word;   // 异常代码
         LastCylceTime : Time;   // 动作时间
         sp : Array[1..16] of Byte;   // 静态变量
      END_STRUCT;
      Status : Struct   // 静态变量
         Busy : Bool;   // Busy
         OkToStart : Bool;   // 静态变量
         NotReadyV2 : Bool;   // 未就绪，请查看故障信息 ！
         TaskDone : Bool;   // 完成
         TaskIO : Bool;   // 合格
         TaskNIO : Bool;   // 失败
         HomePos : Bool;   // 在原点
         PromptValue : Int;   // 提示信息字
      END_STRUCT;
      AtStatus : Word;   // 静态变量
      "Step" : Struct   // 当前运行步
         Main : Int;   // 静态变量
      END_STRUCT;
      CmdMid : Struct   // 命令中间位
         ProgStart : Bool;   // 静态变量
         GoHome : Bool;   // 静态变量
         Stop : Bool;   // 静态变量
      END_STRUCT;
      AtCmdMid : Word;   // 静态变量
      Bus_IN_Data : Struct   // From Input of DP Slave
         AlarmStop : Bool;   // 专用 紧急关断环路关闭（常闭）
         UserSaf : Bool;   // 专用 操作人员防护装置关闭
         Stopmess : Bool;   // 专用 集合故障（常开）
         Alarm_Stop_Intern : Bool;   // 专用 内部紧急关断（常闭）
         Pro_Act : Bool;   // 专用 程序激活
         IN_home : Bool;   // 专用 机器人在原点位置
         On_Path : Bool;   // 专用 机器人在轨迹上
         Robot_Rdy : Bool;   // 专用 机器人控制器就绪
         T1 : Bool;   // 专用 测试1运行
         T2 : Bool;   // 专用 测试2运行
         AUT : Bool;   // 专用 自动运行
         EXT : Bool;   // 专用 外部自动运行
         Peri_Rdy : Bool;   // 专用 驱动装置处于待机运行状态
         Rob_Stopped : Bool;   // 专用 机器人停止
         SP02 : Bool;   // 静态变量
         SP03 : Bool;   // 静态变量
         RecoveryActive : Bool;   // 程序恢复中
         CmdDone : Bool;   // 命令完成
         CmdRdy : Bool;   // 机器人准备好
         ProgReset : Bool;   // 程序复位
         SP04 : Byte;   // 静态变量
         Go_iCmd : Byte;   // 命令反馈（程序号）
         Go_iApplErrNo : Byte;   // 错误代码
         Go_iApplInfNo : Byte;   // 信息提示
         Gp330 : Byte;   // 静态变量
         UserDefineRobOut : Array[8..63] of Byte;   // 静态变量
      END_STRUCT;
      Bus_Out_Data : Struct   // From Input of DP Slave
         Move_Enable : Bool;   // 专用 运行开通
         Ext_Start : Bool;   // 专用外部启动
         Conf_Mess : Bool;   // 专用 错误确认
         Drives_On : Bool;   // 专用 驱动装置接通
         Drives_Off : Bool;   // 专用 驱动装置关闭
         SP01 : Bool;   // 静态变量
         SP02 : Bool;   // 静态变量
         SP03 : Bool;   // 静态变量
         Recovery : Bool;   // 专用 主程序恢复
         Ext_Stop : Bool;   // 专用 外部停止
         AplFaultQuit : Bool;   // 专用 错误清除
         CmdStart : Bool;   // 专用 命令启动
         SP04 : Byte;   // 静态变量
         SP05 : Byte;   // 静态变量
         Gi_iCmd : Byte;   // 专用 命令(程序号)
         Gi_iRobotSpeed : Byte;   // 专用 机器人监控速度
         SP06 : Byte;   // 静态变量
         SP07 : Byte;   // 静态变量
         UserDefineRobIn : Array[8..63] of Byte;   // 用户自定义
      END_STRUCT;
      Info_Err : Struct   // 静态变量
         InfoStruct : Struct   // 信息
            ModeOff : Bool;   // A00. ModeOff !
            OKToStart : Bool;   // A01. OK To Start !
            WaitUserCmdOff : Bool;   // A02.Wait User Command = Off!
            sp03 : Bool;   // A03.
            WaitBusyOff : Bool;   // A04. Wait IO.Busy = Off
            WaitIO_END : Bool;   // A05. Wait IO.END = ON, Check K3
            WaitIO_Move : Bool;   // A06. Wait IO.Move = Off, Check K12=?, K23=Move
            WatiCmdRdy : Bool;   // A07. Wait Cmd Ready!
            WaitChangeProg : Bool;   // A10. Wait Change Prog
            Sp11 : Bool;   // A11.
            Sp12 : Bool;   // A12.
            sp13 : Bool;   // A13.
            StartChangeProg : Bool;   // A14. Start Change Prog
            DriversOn : Bool;   // A15. Start Drivers on!
            Ext_Start : Bool;   // A16.Start Ext Start!
            Recovery : Bool;   // A17.Start Recovery!
            CmdStart : Bool;   // A20.Start CmdStart!
            CmdDone : Bool;   // A21.Wait Done
            xx_5 : Bool;   // A22.
            xx_4 : Bool;   // A23.
            xx_3 : Bool;   // A24.
            xx : Bool;   // A25.
            xx_1 : Bool;   // A26.
            xx_2 : Bool;   // A27.
            xx_10 : Bool;   // A30.
            xx_11 : Bool;   // A31
            xx_12 : Bool;   // A32
            x : Bool;   // A33
            xx_13 : Bool;   // A34
            x_1 : Bool;   // A35
            x_2 : Bool;   // A36
            A37 : Bool;   // A37.
         END_STRUCT;
         ErrStruct : Struct   // 故障
            BusConnectErr : Bool;   // E00. Connnect Err, Pls Reset!
            EndOfTimeOut : Bool;   // E01. Cmd end of time Out !
            AlarmStopErr : Bool;   // E02. Alarm stop!
            UserSafErr : Bool;   // E03. User Saf!
            StopMessErr : Bool;   // E04. Stop mess!
            AlarmStopInternErr : Bool;   // E05.Alarm stop intern!
            T1Mode : Bool;   // E06.in T1 Mode!
            T2Mode : Bool;   // E07.in T2 Mode!
            AutMode : Bool;   // E10.in AUT Mode!
            RobotNotRdy : Bool;   // E11.Robot is not ready!
            Sp12 : Bool;   // E12.
            sp37 : Bool;   // E13.
            sp36 : Bool;   // E14.
            sp35 : Bool;   // E15
            sp34 : Bool;   // E16.
            sp33 : Bool;   // E17.
            sp31 : Bool;   // E20.
            xx_7 : Bool;   // E21.
            xx_6 : Bool;   // E22
            xx_5 : Bool;   // E23
            xx_4 : Bool;   // E24
            xx : Bool;   // E25
            xx_1 : Bool;   // E26
            x : Bool;   // E27
            x_1 : Bool;   // E30
            x_2 : Bool;   // E31
            x_3 : Bool;   // E32
            x_4 : Bool;   // E33
            x_5 : Bool;   // E34
            x_6 : Bool;   // E35
            E36 : Bool;   // E36.
            E37 : Bool;   // E37
         END_STRUCT;
      END_STRUCT;
      AtInfo_Err : Struct   // 静态变量
         Info : DWord;   // 静态变量
         Err : DWord;   // 静态变量
      END_STRUCT;
      FB_Prompt_Object : "FB1022_Prompt_ObjectV2";   // 信息
      Timer_TimeOut : "FB951_SDTimerV2";   // 完成超时
      TimdDrivers_Off : "FB951_SDTimerV2";   // 静态变量
      Stack : Struct   // 静态变量
         Index : Int;   // 静态变量
         "Step" : Array[0..9] of Int;   // 最高允许10级嵌套
         sp : Array[0..1] of Int;   // 静态变量
      END_STRUCT;
      Aux : Struct   // 静态变量
         JpEnd : Bool;   // 静态变量
         ReqPosContinuous : Bool;   // 静态变量
         DPRD_RetVal : Int;   // 静态变量
         DPWR_RetVal : Int;   // 静态变量
         RetVal : Int;   // 静态变量
         Index : Int;   // 静态变量
         timStart : Time;   // 静态变量
         T_Prog : Byte;   // 静态变量
         sp : Array[0..100] of Byte;   // 静态变量
      END_STRUCT;
      lastAddr : Int := 398;   // 静态变量
      CycleTime : Int;   // 静态变量
      PromptValueBake : Int;   // 静态变量
      ShiftBake : Int;   // 静态变量
      StartTime : Time;   // 静态变量
      ET : Time;   // 静态变量
      IN_EDGE : Bool;   // 静态变量
   END_VAR
   VAR_TEMP
      AnyCmdOn : Bool;   // 临时变量
      T_bNextStep_ThisCycle : Bool;   // 下一步，返回再次扫描Case的下一步程序
      T_DWORD : DWord;   // 临时变量
      T_Dint : DInt;   // 临时变量
      T_Word : Word;   // 临时变量
      T_int : Int;   // 临时变量
      T_int2 : Int;   // 临时变量
      T_Byte : Int;   // 临时变量
      T_RetVal : Int;   // 临时变量
   END_VAR
   VAR CONSTANT
      STEP_EndScan : Int := 28000;   // 最终执行的程序步,100%扫描
      OK : Int := 1;
      JP1 : Int := 2;
      JP2 : Int := 3;
      JP3 : Int := 4;
   END_VAR
BEGIN

   // ---------- 网络 1 ----------
   // 含义：本网络为 StructuredText（SCL）原文重建，非 LAD 折叠
   IF TRUE THEN
       IF #ManMode = false
       THEN
           #TP_Cmd := 0;
       END_IF;
       #AtCmdMid := #TP_Cmd OR #AtCmd.Auto;
       IF #AtCmdMid <> 0
       THEN
           #AnyCmdOn := true;
       ELSE
           #AnyCmdOn := false;
           IF #Status.Busy = FALSE AND
               #ErrRst = FALSE AND
               #AllMode = TRUE
           THEN
               "FC1003_CR"(Jp => #Aux.JpEnd);
               IF #Aux.JpEnd = TRUE
               THEN
                   RETURN;
               END_IF;
           END_IF;
       END_IF;
       #TP_Status := #AtStatus;
   END_IF;
   IF TRUE THEN
       #Aux.DPRD_RetVal := DPRD_DAT(LADDR := #CTRL_IN.InitParameter.HW_Addr, RECORD => #Bus_IN_Data);
       #Status.HomePos := #Bus_IN_Data.IN_home;
       #CTRL_OUT.ProgNo := #Bus_IN_Data.Go_iCmd;
       IF (#EMMode = false) AND
           (#RobotEnble = TRUE)
       THEN
           #Bus_Out_Data.Move_Enable := TRUE;
       ELSE
           #Bus_Out_Data.Move_Enable := false;
       END_IF;
       #TimdDrivers_Off();
       #TimdDrivers_Off.IN := #Bus_Out_Data.Move_Enable;
       #TimdDrivers_Off.TV := T#0.6S;
       #Bus_Out_Data.Drives_Off := #TimdDrivers_Off.Q;
   END_IF;
   IF TRUE THEN
       IF #Info_Err.ErrStruct.BusConnectErr = FALSE AND
           #Bus_IN_Data.EXT = TRUE AND
           #Bus_IN_Data.Robot_Rdy = TRUE AND
           #Bus_IN_Data.Go_iApplErrNo = 0
       THEN
           #Status.OkToStart := TRUE;
       ELSE
           #Status.OkToStart := FALSE;
       END_IF;
       IF #Status.OkToStart = FALSE
       THEN
           #Status.NotReadyV2 := TRUE;
       ELSE
           #Status.NotReadyV2 := FALSE;
       END_IF;
   END_IF;
   IF TRUE THEN
       #Info_Err.InfoStruct.ModeOff := NOT (#AllMode);
       #Info_Err.InfoStruct.OKToStart := #Status.OkToStart AND (NOT (#Status.Busy));
       #Info_Err.InfoStruct.Ext_Start := #Bus_Out_Data.Ext_Start;
       #Info_Err.InfoStruct.Recovery := #Bus_Out_Data.Recovery;
       #Info_Err.InfoStruct.CmdStart := #Bus_Out_Data.CmdStart;
       #Info_Err.InfoStruct.CmdDone := #Bus_IN_Data.CmdDone;
   END_IF;
   IF TRUE THEN
       IF #Aux.DPRD_RetVal <> 0
       THEN
           #Aux.ReqPosContinuous := FALSE;
           #Info_Err.ErrStruct.BusConnectErr := true;
       ELSE
           #Info_Err.ErrStruct.BusConnectErr := false;
           #Info_Err.ErrStruct.AlarmStopErr := NOT (#Bus_IN_Data.AlarmStop);
           #Info_Err.ErrStruct.UserSafErr := NOT (#Bus_IN_Data.UserSaf);
           #Info_Err.ErrStruct.StopMessErr := (#Bus_IN_Data.Stopmess);
           #Info_Err.ErrStruct.AlarmStopInternErr := NOT (#Bus_IN_Data.Alarm_Stop_Intern);
           #Info_Err.ErrStruct.T1Mode := (#Bus_IN_Data.T1);
           #Info_Err.ErrStruct.T2Mode := (#Bus_IN_Data.T2);
           #Info_Err.ErrStruct.AutMode := (#Bus_IN_Data.AUT);
           #Info_Err.ErrStruct.RobotNotRdy := NOT (#Bus_IN_Data.Robot_Rdy);
           #CTRL_OUT.ErrorCode := #Bus_IN_Data.Go_iApplErrNo;
       END_IF;
   END_IF;
   IF TRUE THEN
       IF (#ErrRst = TRUE OR
           (#AnyCmdOn = TRUE AND #Status.OkToStart = TRUE))
           AND
           #Status.Busy = FALSE AND
           #AllMode = TRUE
       THEN
           #Status.Busy := true;
           #AtInfo_Err.Info := 0;
           #AtInfo_Err.Err := 0;
           #Timer_TimeOut.IN := FALSE;
           #Timer_TimeOut.TV := #CTRL_IN.InitParameter.TimeOutSetValue;
           #Step.Main := 1;
       END_IF;
       IF #Status.Busy = TRUE
       THEN
           IF "Debug_True" = FALSE
           THEN
               #Info_Err.ErrStruct.EndOfTimeOut := #Timer_TimeOut.Q;
           END_IF;
           IF #AllMode = FALSE OR
               #Info_Err.ErrStruct.EndOfTimeOut OR
               #Cmd.Auto.Stop = TRUE
           THEN
               IF #Step.Main < #STEP_EndScan THEN
                   #Step.Main := #STEP_EndScan;
               END_IF;
           END_IF;
           #Timer_TimeOut();
           IF #Timer_TimeOut.IN = TRUE
           THEN
               #CTRL_OUT.LastCylceTime := #Timer_TimeOut.ET;
           END_IF;
       END_IF;
   END_IF;
   IF TRUE THEN
       #T_bNextStep_ThisCycle := FALSE;
   _Scan_Case:
       ;

       CASE #Step.Main OF
           1:
               IF TRUE
               THEN
                   #Status.TaskIO := FALSE;
                   #Status.TaskNIO := FALSE;
                   #Stack.Index := 0;
                   #Timer_TimeOut.IN := TRUE;
                   IF #AnyCmdOn = true
                   THEN
                       IF (#Bus_IN_Data.Robot_Rdy = FALSE OR
                           #Bus_IN_Data.Go_iApplErrNo <> 0)
                       THEN
                           #Bus_Out_Data.Conf_Mess := TRUE;
                           #Bus_Out_Data.AplFaultQuit := true;
                           IF (#Bus_IN_Data.Go_iApplErrNo <> 0)
                           THEN
                               #Bus_Out_Data.Recovery := TRUE;
                           END_IF;
                       ELSE
                           #Bus_Out_Data.Conf_Mess := FALSE;
                           #Bus_Out_Data.AplFaultQuit := false;
                           #Bus_Out_Data.Recovery := FALSE;
                           IF (TRUE)
                           THEN
                               #Step.Main := (ENCO(IN := SWAP(IN := #AtCmdMid)) + 1) * 1000;
                               #T_bNextStep_ThisCycle := true;
                           END_IF;
                       END_IF;
                   ELSE
                       IF (#Bus_IN_Data.Robot_Rdy = FALSE OR
                           #Bus_IN_Data.Go_iApplErrNo <> 0) AND
                           (#Bus_IN_Data.EXT)
                       THEN
                           #Bus_Out_Data.Conf_Mess := TRUE;
                           #Bus_Out_Data.AplFaultQuit := true;
                           IF (#Bus_IN_Data.Go_iApplErrNo <> 0)
                           THEN
                               #Bus_Out_Data.Recovery := TRUE;
                           END_IF;
                       ELSE
                           #Bus_Out_Data.Conf_Mess := FALSE;
                           #Bus_Out_Data.AplFaultQuit := false;
                           #Status.TaskIO := true;
                           #Bus_Out_Data.Recovery := FALSE;
                           #Step.Main := #STEP_EndScan;
                       END_IF;
                   END_IF;
                   #Aux.ReqPosContinuous := FALSE;
               END_IF;
           1001:
               IF TRUE
               THEN
                   #Aux.T_Prog := #CTRL_IN.ProgNo;
                   IF (#Bus_IN_Data.Peri_Rdy = TRUE) AND
                       (#Bus_IN_Data.Pro_Act = TRUE)
                   THEN
                       #Step.Main := 1006;
                   ELSE
                       IF (#Bus_Out_Data.Drives_Off = false)
                       THEN
                           #Step.Main := 1002;
                       ELSE
                           #TimdDrivers_Off.IN := FALSE;
                       END_IF;
                   END_IF;
               END_IF;
           1002:
               IF (#Bus_Out_Data.Drives_Off = TRUE)
               THEN
                   #T_bNextStep_ThisCycle := TRUE;
               END_IF;
           1003:
               IF (#Bus_IN_Data.Peri_Rdy = TRUE)
               THEN
                   #Bus_Out_Data.Drives_On := false;
                   #T_bNextStep_ThisCycle := true;
               ELSE
                   #Bus_Out_Data.Drives_On := TRUE;
               END_IF;
           1004:
               IF (#Bus_IN_Data.EXT = TRUE)
               THEN
                   #Bus_Out_Data.Ext_Start := FALSE;
                   #T_bNextStep_ThisCycle := true;
               ELSE
                   #Bus_Out_Data.Ext_Start := true;
               END_IF;
           1005:
               IF (#Bus_IN_Data.RecoveryActive = true)
               THEN
                   #Bus_Out_Data.Recovery := false;
                   #T_bNextStep_ThisCycle := true;
               ELSE
                   #Bus_Out_Data.Recovery := true;
               END_IF;
           1006:
               #Bus_Out_Data.Gi_iCmd := #Aux.T_Prog;
               IF (#Bus_IN_Data.Peri_Rdy = true) AND
                   (#Bus_IN_Data.Pro_Act = true)
               THEN
                   #T_bNextStep_ThisCycle := true;
               END_IF;
           1007:
               IF (#Bus_IN_Data.Go_iCmd = #Aux.T_Prog)
               THEN
                   #T_bNextStep_ThisCycle := true;
                   #Info_Err.InfoStruct.WaitChangeProg := FALSE;
               ELSE
                   #Bus_Out_Data.Gi_iCmd := #Aux.T_Prog;
                   #Info_Err.InfoStruct.WaitChangeProg := FALSE;
               END_IF;
           1008:
               IF #Bus_IN_Data.CmdRdy
               THEN
                   #T_bNextStep_ThisCycle := true;
                   #Info_Err.InfoStruct.WatiCmdRdy := FALSE;
               ELSE
                   #Info_Err.InfoStruct.WatiCmdRdy := TRUE;
               END_IF;
           1009:
               IF #Bus_IN_Data.CmdDone
               THEN
                   #Bus_Out_Data.CmdStart := FALSE;
                   #T_bNextStep_ThisCycle := true;
               ELSE
                   #Bus_Out_Data.CmdStart := TRUE;
               END_IF;
           1010:
               IF #Bus_IN_Data.CmdRdy = true
               THEN
                   #Status.TaskIO := true;
                   #T_bNextStep_ThisCycle := true;
               END_IF;
           2001:
               IF TRUE
               THEN
                   #CTRL_IN.ProgNo := 255;
                   #Aux.T_Prog := #CTRL_IN.ProgNo;
                   IF (#Bus_IN_Data.Peri_Rdy = TRUE) AND
                       (#Bus_IN_Data.Pro_Act = TRUE)
                   THEN
                       #Step.Main := 1007;
                   ELSE
                       IF (#Bus_Out_Data.Drives_Off = false)
                       THEN
                           #Step.Main := 1002;
                       ELSE
                           #TimdDrivers_Off.IN := FALSE;
                       END_IF;
                   END_IF;
               END_IF;
           3001:
               #Bus_Out_Data.Ext_Stop := TRUE;
               #T_bNextStep_ThisCycle := true;
           1011, 3002:
               IF TRUE
               THEN
                   IF #Stack.Index >= 1
                   THEN
                       #Stack.Index := #Stack.Index - 1;
                       #Step.Main := #Stack.Step[#Stack.Index];
                   ELSE
                       #Status.TaskDone := true;
                       #Step.Main := #STEP_EndScan;
                   END_IF;
               END_IF;
           #STEP_EndScan:
               IF (#Bus_IN_Data.Rob_Stopped = TRUE)
               THEN
                   #Bus_Out_Data.Ext_Stop := FALSE;
                   #T_bNextStep_ThisCycle := true;
               ELSE
                   #Bus_Out_Data.Ext_Stop := TRUE;
               END_IF;
           28001:
               IF (#Bus_IN_Data.CmdRdy = FALSE)
               THEN
                   #T_bNextStep_ThisCycle := true;
               ELSE
                   #Step.Main := 28003;
               END_IF;
           28002:
               IF (#Bus_IN_Data.Pro_Act = FALSE)
               THEN
                   #T_bNextStep_ThisCycle := true;
                   #Bus_Out_Data.Ext_Stop := FALSE;
               ELSE
                   #Bus_Out_Data.Ext_Stop := TRUE;
               END_IF;
           28003:
               #Timer_TimeOut.IN := FALSE;
               #Bus_Out_Data.Drives_On := FALSE;
               #Bus_Out_Data.Ext_Start := FALSE;
               #Bus_Out_Data.Recovery := FALSE;
               #Bus_Out_Data.CmdStart := FALSE;
               #Bus_Out_Data.Ext_Stop := FALSE;
               #Bus_Out_Data.AplFaultQuit := FALSE;
               #Bus_Out_Data.Conf_Mess := FALSE;
               #Timer_TimeOut.IN := FALSE;
               #Status.TaskDone := TRUE;
               IF #Status.TaskIO = FALSE
               THEN
                   #Status.TaskNIO := true;
               ELSE
                   #Status.TaskNIO := FALSE;
               END_IF;
               IF #AnyCmdOn = false
               THEN
                   #Status.TaskDone := false;
                   #Info_Err.InfoStruct.WaitUserCmdOff := false;
                   #T_bNextStep_ThisCycle := true;
               ELSE
                   #AtCmd.Auto := 0;
                   #Info_Err.InfoStruct.WaitUserCmdOff := true;
               END_IF;
           28004:
               IF TRUE
               THEN
                   #Status.Busy := FALSE;
                   #Step.Main := 0;
               END_IF;
           ELSE
               ;
       END_CASE;
       IF #T_bNextStep_ThisCycle = TRUE
       THEN
           #Step.Main := #Step.Main + 1;
           GOTO _Scan_Case;
       END_IF;
   END_IF;
   IF TRUE THEN
       IF #AllMode = FALSE
       THEN
           ;
       END_IF;
       IF TRUE THEN
           #Aux.DPWR_RetVal := DPWR_DAT(LADDR := #CTRL_IN.InitParameter.HW_Addr, RECORD := #Bus_Out_Data);
       END_IF;
       IF TRUE
       THEN
           ;
       END_IF;
   END_IF;
   IF TRUE THEN
       IF "DB1000_StdSignal".PLS.PS10
       THEN
           #Status.PromptValue := #FB_Prompt_Object.PromptValue;
       END_IF;
   END_IF;
   IF "DB1060_AutoStep".HorDrillAutoStep.HorDrillStep.StepStart OR
       "DB1060_AutoStep".DownDrillAutoStep.DownDrillStep.StepStart OR
       "DB720_KuKa_MainCtrl".CheckBit.StepStart OR
       "DB720_KuKa_MainCtrl".ChangeTool.StepStart OR
       "DB1060_AutoStep".DiamondAutoStep.DiamondStep.StepStart
   THEN
       #Bus_Out_Data.Gi_iRobotSpeed := #CTRL_IN.RobotSpeed;
   ELSE
       #Bus_Out_Data.Gi_iRobotSpeed := 30;
   END_IF;
END_FUNCTION_BLOCK

FUNCTION "FC1900_Communication_PC" : Void   // FC1900, LAD
{ S7_Optimized_Access := 'TRUE' }
VERSION : 0.1
   VAR_TEMP
      Angle : DInt;
      width : DInt;
      SwingSpeed : DInt;
   END_VAR
BEGIN

REGION Network 1: 机器人回原点
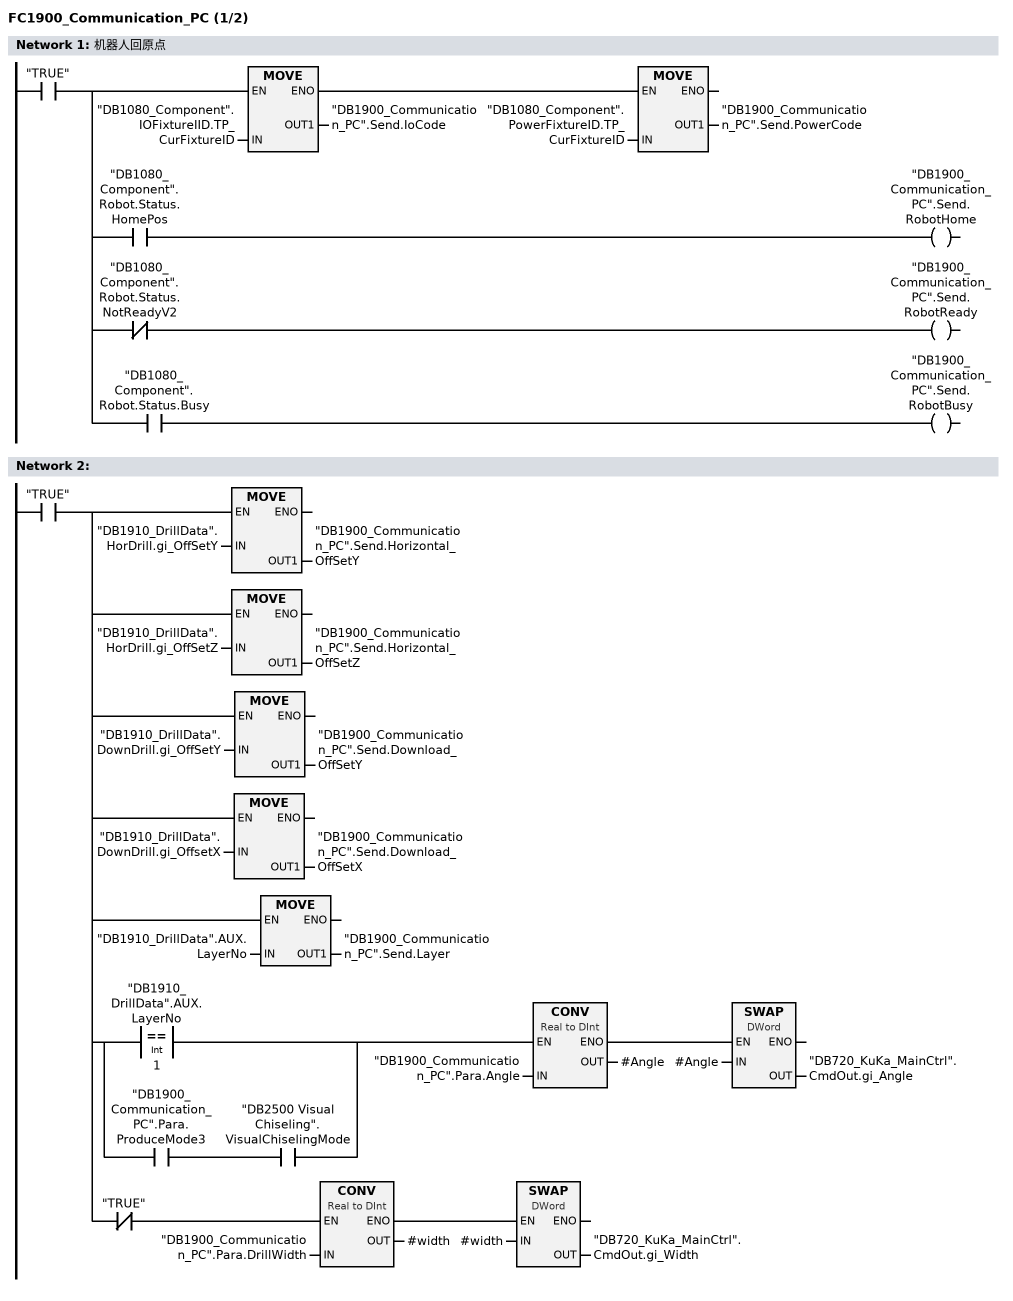
   RUNG wire#powerrail
      Contact( "TRUE" )
      wire#w1
      Move(in := "DB1080_Component".IOFixtureIID.TP_CurFixtureID, out1 => "DB1900_Communication_PC".Send.IoCode)
      Move(in := "DB1080_Component".PowerFixtureID.TP_CurFixtureID, out1 => "DB1900_Communication_PC".Send.PowerCode)
   END_RUNG
   RUNG wire#w1
      Contact( "DB1080_Component".Robot.Status.HomePos )
      Coil( "DB1900_Communication_PC".Send.RobotHome )
   END_RUNG
   RUNG wire#w1
      I_Contact( "DB1080_Component".Robot.Status.NotReadyV2 )
      Coil( "DB1900_Communication_PC".Send.RobotReady )
   END_RUNG
   RUNG wire#w1
      Contact( "DB1080_Component".Robot.Status.Busy )
      Coil( "DB1900_Communication_PC".Send.RobotBusy )
   END_RUNG
   // the same network as SCL:
   IF "TRUE" THEN
       "DB1900_Communication_PC".Send.IoCode := "DB1080_Component".IOFixtureIID.TP_CurFixtureID;
       "DB1900_Communication_PC".Send.PowerCode := "DB1080_Component".PowerFixtureID.TP_CurFixtureID;
   END_IF;
   "DB1900_Communication_PC".Send.RobotHome := "TRUE" AND "DB1080_Component".Robot.Status.HomePos;
   "DB1900_Communication_PC".Send.RobotReady := "TRUE" AND NOT "DB1080_Component".Robot.Status.NotReadyV2;
   "DB1900_Communication_PC".Send.RobotBusy := "TRUE" AND "DB1080_Component".Robot.Status.Busy;
END_REGION

REGION Network 2
   IF "TRUE" THEN
       "DB1900_Communication_PC".Send.Horizontal_OffSetY := "DB1910_DrillData".HorDrill.gi_OffSetY;
       "DB1900_Communication_PC".Send.Horizontal_OffSetZ := "DB1910_DrillData".HorDrill.gi_OffSetZ;
       "DB1900_Communication_PC".Send.Download_OffSetY := "DB1910_DrillData".DownDrill.gi_OffSetY;
       "DB1900_Communication_PC".Send.Download_OffSetX := "DB1910_DrillData".DownDrill.gi_OffsetX;
       "DB1900_Communication_PC".Send.Layer := "DB1910_DrillData".AUX.LayerNo;
   END_IF;
   IF "TRUE" AND (("DB1910_DrillData".AUX.LayerNo = 1) OR ("DB1900_Communication_PC".Para.ProduceMode3 AND "DB2500 Visual Chiseling".VisualChiselingMode)) THEN
       #Angle := REAL_TO_DINT("DB1900_Communication_PC".Para.Angle);
       "DB720_KuKa_MainCtrl".CmdOut.gi_Angle := SWAP(#Angle);
   END_IF;
   IF "TRUE" AND NOT "TRUE" THEN
       #width := REAL_TO_DINT("DB1900_Communication_PC".Para.DrillWidth);
       "DB720_KuKa_MainCtrl".CmdOut.gi_Width := SWAP(#width);
   END_IF;
END_REGION

REGION Network 3: 角度设置超限！
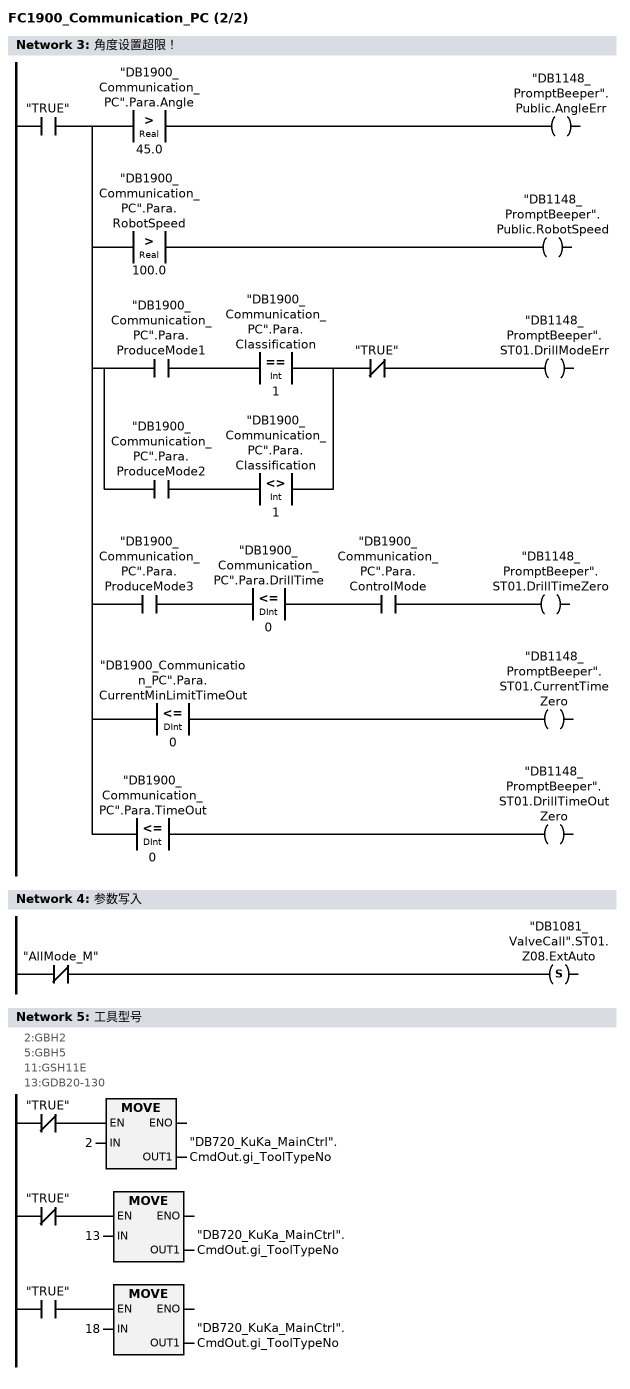
   RUNG wire#powerrail
      Contact( "TRUE" )
      wire#w1
      { S7_Templates := "SrcType := Real" } GT_Contact(in1 := "DB1900_Communication_PC".Para.Angle, in2 := 45.0)
      Coil( "DB1148_PromptBeeper".Public.AngleErr )
   END_RUNG
   RUNG wire#w1
      { S7_Templates := "SrcType := Real" } GT_Contact(in1 := "DB1900_Communication_PC".Para.RobotSpeed, in2 := 100.0)
      Coil( "DB1148_PromptBeeper".Public.RobotSpeed )
   END_RUNG
   RUNG wire#w1
      Contact( "DB1900_Communication_PC".Para.ProduceMode1 )
      { S7_Templates := "SrcType := Int" } EQ_Contact(in1 := "DB1900_Communication_PC".Para.Classification, in2 := 1)
      wire#w2
      I_Contact( "TRUE" )
      Coil( "DB1148_PromptBeeper".ST01.DrillModeErr )
   END_RUNG
   RUNG wire#w1
      Contact( "DB1900_Communication_PC".Para.ProduceMode2 )
      { S7_Templates := "SrcType := Int" } NE_Contact(in1 := "DB1900_Communication_PC".Para.Classification, in2 := 1)
   END_RUNG wire#w2
   RUNG wire#w1
      Contact( "DB1900_Communication_PC".Para.ProduceMode3 )
      { S7_Templates := "SrcType := DInt" } LE_Contact(in1 := "DB1900_Communication_PC".Para.DrillTime, in2 := 0)
      Contact( "DB1900_Communication_PC".Para.ControlMode )
      Coil( "DB1148_PromptBeeper".ST01.DrillTimeZero )
   END_RUNG
   RUNG wire#w1
      { S7_Templates := "SrcType := DInt" } LE_Contact(in1 := "DB1900_Communication_PC".Para.CurrentMinLimitTimeOut, in2 := 0)
      Coil( "DB1148_PromptBeeper".ST01.CurrentTimeZero )
   END_RUNG
   RUNG wire#w1
      { S7_Templates := "SrcType := DInt" } LE_Contact(in1 := "DB1900_Communication_PC".Para.TimeOut, in2 := 0)
      Coil( "DB1148_PromptBeeper".ST01.DrillTimeOutZero )
   END_RUNG
   // the same network as SCL:
   "DB1148_PromptBeeper".Public.AngleErr := "TRUE" AND ("DB1900_Communication_PC".Para.Angle > 45.0);
   "DB1148_PromptBeeper".Public.RobotSpeed := "TRUE" AND ("DB1900_Communication_PC".Para.RobotSpeed > 100.0);
   "DB1148_PromptBeeper".ST01.DrillModeErr := "TRUE" AND (("DB1900_Communication_PC".Para.ProduceMode1 AND ("DB1900_Communication_PC".Para.Classification = 1)) OR ("DB1900_Communication_PC".Para.ProduceMode2 AND ("DB1900_Communication_PC".Para.Classification <> 1))) AND NOT "TRUE";
   "DB1148_PromptBeeper".ST01.DrillTimeZero := "TRUE" AND "DB1900_Communication_PC".Para.ProduceMode3 AND ("DB1900_Communication_PC".Para.DrillTime <= 0) AND "DB1900_Communication_PC".Para.ControlMode;
   "DB1148_PromptBeeper".ST01.CurrentTimeZero := "TRUE" AND ("DB1900_Communication_PC".Para.CurrentMinLimitTimeOut <= 0);
   "DB1148_PromptBeeper".ST01.DrillTimeOutZero := "TRUE" AND ("DB1900_Communication_PC".Para.TimeOut <= 0);
END_REGION

REGION Network 4: 参数写入
   RUNG wire#powerrail
      I_Contact( "AllMode_M" )
      S_Coil( "DB1081_ValveCall".ST01.Z08.ExtAuto )
   END_RUNG
   // the same network as SCL:
   IF NOT "AllMode_M" THEN "DB1081_ValveCall".ST01.Z08.ExtAuto := TRUE; END_IF;
END_REGION

REGION Network 5: 工具型号
   // 2:GBH2
   // 5:GBH5
   // 11:GSH11E
   // 13:GDB20-130
   RUNG wire#powerrail
      I_Contact( "TRUE" )
      Move(in := 2, out1 => "DB720_KuKa_MainCtrl".CmdOut.gi_ToolTypeNo)
   END_RUNG
   RUNG wire#powerrail
      I_Contact( "TRUE" )
      Move(in := 13, out1 => "DB720_KuKa_MainCtrl".CmdOut.gi_ToolTypeNo)
   END_RUNG
   RUNG wire#powerrail
      Contact( "TRUE" )
      Move(in := 18, out1 => "DB720_KuKa_MainCtrl".CmdOut.gi_ToolTypeNo)
   END_RUNG
   // the same network as SCL:
   IF NOT "TRUE" THEN
       "DB720_KuKa_MainCtrl".CmdOut.gi_ToolTypeNo := 2;
       "DB720_KuKa_MainCtrl".CmdOut.gi_ToolTypeNo := 13;
   END_IF;
   IF "TRUE" THEN "DB720_KuKa_MainCtrl".CmdOut.gi_ToolTypeNo := 18; END_IF;
END_REGION
END_FUNCTION

// folder: 005_Component/Cooling Fan

FUNCTION_BLOCK "FB2008_CoolingFan"   // FB2008, SCL
{ S7_Optimized_Access := 'TRUE' }
// ============================================================
//  Block: FB2008_CoolingFan
//  ============================================================
//  编号：FB2008
//  原始语言：LAD（规则翻译为 SCL）
//  含义：由 LAD/FBD 网络折叠生成的等效 SCL，导入前请人工复核
   VAR_INPUT
      Man_Mode : Bool;   // 输入参数
      Auto_Mode : Bool;   // 输入参数
      Emm_Mode : Bool;   // 输入参数
      I_StationToolOn_1 : Bool;   // 输入参数
      I_StationToolOn_2 : Bool;   // 输入参数
      CoolingTime : Time;   // 输入参数
   END_VAR
   VAR_OUTPUT
      Q_StationCoolingFan : Bool;   // 输出参数
   END_VAR
   VAR
      "A Station CoolingFan" : "FB2009_CoolingFanFunction";   // 静态变量
      "B Station CoolingFan" : "FB2009_CoolingFanFunction";   // 静态变量
      "C Station CoolingFan" : "FB2009_CoolingFanFunction";   // 静态变量
      SR_StationTool : Bool;   // 静态变量
      ToolAtPos : Bool;   // 静态变量
      Timer_StationToolOn : IEC_TIMER;   // 静态变量
      Timer_StationCoolingFan : IEC_TIMER;   // 静态变量
      PT : Time;   // 静态变量
      ET : Time;   // 静态变量
      IN : Bool;   // 静态变量
      Q : Bool;   // 静态变量
   END_VAR
BEGIN

   // ---------- 网络 1 ----------
   // 含义：调用块/实例 #A Station CoolingFan，参数：Man_Mode := "ManMode_M", Auto_Mode := "AutoMode_M", Emm_Mode := "EMMode_M", I_StationToolOn_1 := "AStation_ToolOn1", I_StationToolOn_2 := "AStation_ToolOn2", CoolingTime := T#30M, Q_StationCoolingFan => "QAStationFan"
   #"A Station CoolingFan"(Man_Mode := "ManMode_M",
                           Auto_Mode := "AutoMode_M",
                           Emm_Mode := "EMMode_M",
                           I_StationToolOn_1 := "AStation_ToolOn1",
                           I_StationToolOn_2 := "AStation_ToolOn2",
                           CoolingTime := T#30M,
                           Q_StationCoolingFan => "QAStationFan");

   // ---------- 网络 2 ----------
   // 含义：调用块/实例 #B Station CoolingFan，参数：Man_Mode := "ManMode_M", Auto_Mode := "AutoMode_M", Emm_Mode := "EMMode_M", I_StationToolOn_1 := "BStation_ToolOn1", I_StationToolOn_2 := "BStation_ToolOn2", CoolingTime := T#30M, Q_StationCoolingFan => "QBStationFan"
   #"B Station CoolingFan"(Man_Mode := "ManMode_M",
                           Auto_Mode := "AutoMode_M",
                           Emm_Mode := "EMMode_M",
                           I_StationToolOn_1 := "BStation_ToolOn1",
                           I_StationToolOn_2 := "BStation_ToolOn2",
                           CoolingTime := T#30M,
                           Q_StationCoolingFan => "QBStationFan");

   // ---------- 网络 3 ----------
   // 含义：调用块/实例 #C Station CoolingFan，参数：Man_Mode := "ManMode_M", Auto_Mode := "AutoMode_M", Emm_Mode := "EMMode_M", CoolingTime := T#30M, Q_StationCoolingFan => "QCStationFan"
   #"C Station CoolingFan"(Man_Mode := "ManMode_M",
                           Auto_Mode := "AutoMode_M",
                           Emm_Mode := "EMMode_M",
                           I_StationToolOn_1 := FALSE,
                           I_StationToolOn_2 := FALSE,
                           CoolingTime := T#30M,
                           Q_StationCoolingFan => "QCStationFan");

   // ---------- 网络 4 ----------
   // （空白网络）
END_FUNCTION_BLOCK

FUNCTION_BLOCK "FB2009_CoolingFanFunction"   // FB2009, SCL
{ S7_Optimized_Access := 'TRUE' }
// ============================================================
//  Block: FB2009_CoolingFanFunction
//  ============================================================
//  编号：FB2009
//  原始语言：LAD（规则翻译为 SCL）
//  含义：由 LAD/FBD 网络折叠生成的等效 SCL，导入前请人工复核
   VAR_INPUT
      Man_Mode : Bool;   // 手动模式
      Auto_Mode : Bool;   // 自动模式
      Emm_Mode : Bool;   // 紧急停止模式
      I_StationToolOn_1 : Bool;   // 夹具在位信号1
      I_StationToolOn_2 : Bool;   // 夹具在位信号2
      CoolingTime : Time;   // 冷却时间
   END_VAR
   VAR_OUTPUT
      Q_StationCoolingFan : Bool;   // 散热风扇打开
   END_VAR
   VAR
      SR_StationTool : Bool;   // 静态变量
      ToolAtPos : Bool;   // 工具在位
      Timer_StationToolOn : IEC_TIMER;   // 工具在位接通延时检测
      Timer_StationCoolingFan : IEC_TIMER;   // 风扇冷却接通延时
   END_VAR
BEGIN

   // ---------- 网络 1 ----------
   // 标题：工具在位检测
   // 含义：调用定时器实例 #Timer_StationToolOn.TON
   #Timer_StationToolOn.TON(IN := (#Auto_Mode AND #I_StationToolOn_1) AND #I_StationToolOn_2,
                            PT := T#2s);
   IF (NOT (#I_StationToolOn_1) OR NOT (#I_StationToolOn_2) OR #Timer_StationCoolingFan.Q OR #Man_Mode OR #Emm_Mode) THEN
       #SR_StationTool := FALSE;
   ELSIF #Timer_StationToolOn.Q THEN
       #SR_StationTool := TRUE;
   END_IF;
   #ToolAtPos := #SR_StationTool;
   #Timer_StationCoolingFan.TON(IN := #SR_StationTool,
                                PT := #CoolingTime);

   // ---------- 网络 2 ----------
   // 标题：散热风扇打开
   // 含义：将 #ToolAtPos AND NOT (#Timer_StationCoolingFan.Q) 赋给 #Q_StationCoolingFan
   #Q_StationCoolingFan := #ToolAtPos AND NOT (#Timer_StationCoolingFan.Q);

   // ---------- 网络 3 ----------
   // （空白网络）
END_FUNCTION_BLOCK

// folder: 006_ Visual Chiseling

FUNCTION "FC2100 Modbus TCP" : Void   // FC2100, LAD
TITLE = Communication Program Between PLC and ROS
{ S7_Optimized_Access := 'TRUE' }
VERSION : 0.1
// Programmed by Wang Xinyang, 20220610. Any Problem Please Contact Mr.Wang.
   VAR_TEMP
      High : Bool;
      Low : Bool;
   END_VAR
BEGIN

REGION Network 1: Always 1 and 0
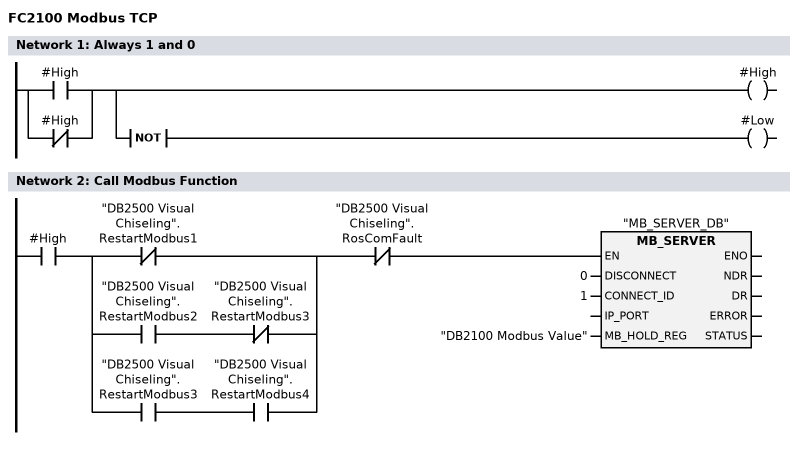
   RUNG wire#powerrail
      Contact( #High )
      wire#w1
      Coil( #High )
   END_RUNG
   RUNG wire#powerrail
      I_Contact( #High )
   END_RUNG wire#w1
   RUNG wire#w1
      Not()
      Coil( #Low )
   END_RUNG
   // the same network as SCL:
   #High := #High OR NOT #High;
   #Low := NOT #High;
END_REGION

REGION Network 2: Call Modbus Function
   IF #High AND (NOT "DB2500 Visual Chiseling".RestartModbus1 OR ("DB2500 Visual Chiseling".RestartModbus2 AND NOT "DB2500 Visual Chiseling".RestartModbus3) OR ("DB2500 Visual Chiseling".RestartModbus3 AND "DB2500 Visual Chiseling".RestartModbus4)) AND NOT "DB2500 Visual Chiseling".RosComFault THEN
       "MB_SERVER_DB"(DISCONNECT := 0, CONNECT_ID := 1, MB_HOLD_REG := "DB2100 Modbus Value");   // MB_SERVER
   END_IF;
END_REGION
END_FUNCTION

FUNCTION "FC2300 Time Calculation" : Void   // FC2300, LAD
TITLE = PLC Transfer Value to ROS
{ S7_Optimized_Access := 'TRUE' }
VERSION : 0.1
// Programmed by Wang Xinyang, 20220610. Any Problem Please Contact Mr.Wang.
   VAR_TEMP
      High : Bool;
      Low : Bool;
      Temp_PLC_Year : UInt;
      Temp_PLC_Month : UInt;
      Temp_PLC_Minute : UInt;
      Temp_ROS_Year : UInt;
      Temp_ROS_MonthDay : UInt;
      Temp_ROS_Month : UInt;
      Temp_ROS_Minute : UInt;
      Temp_PLCRetValue : UInt;
   END_VAR
BEGIN

REGION Network 1: Always 1 and 0
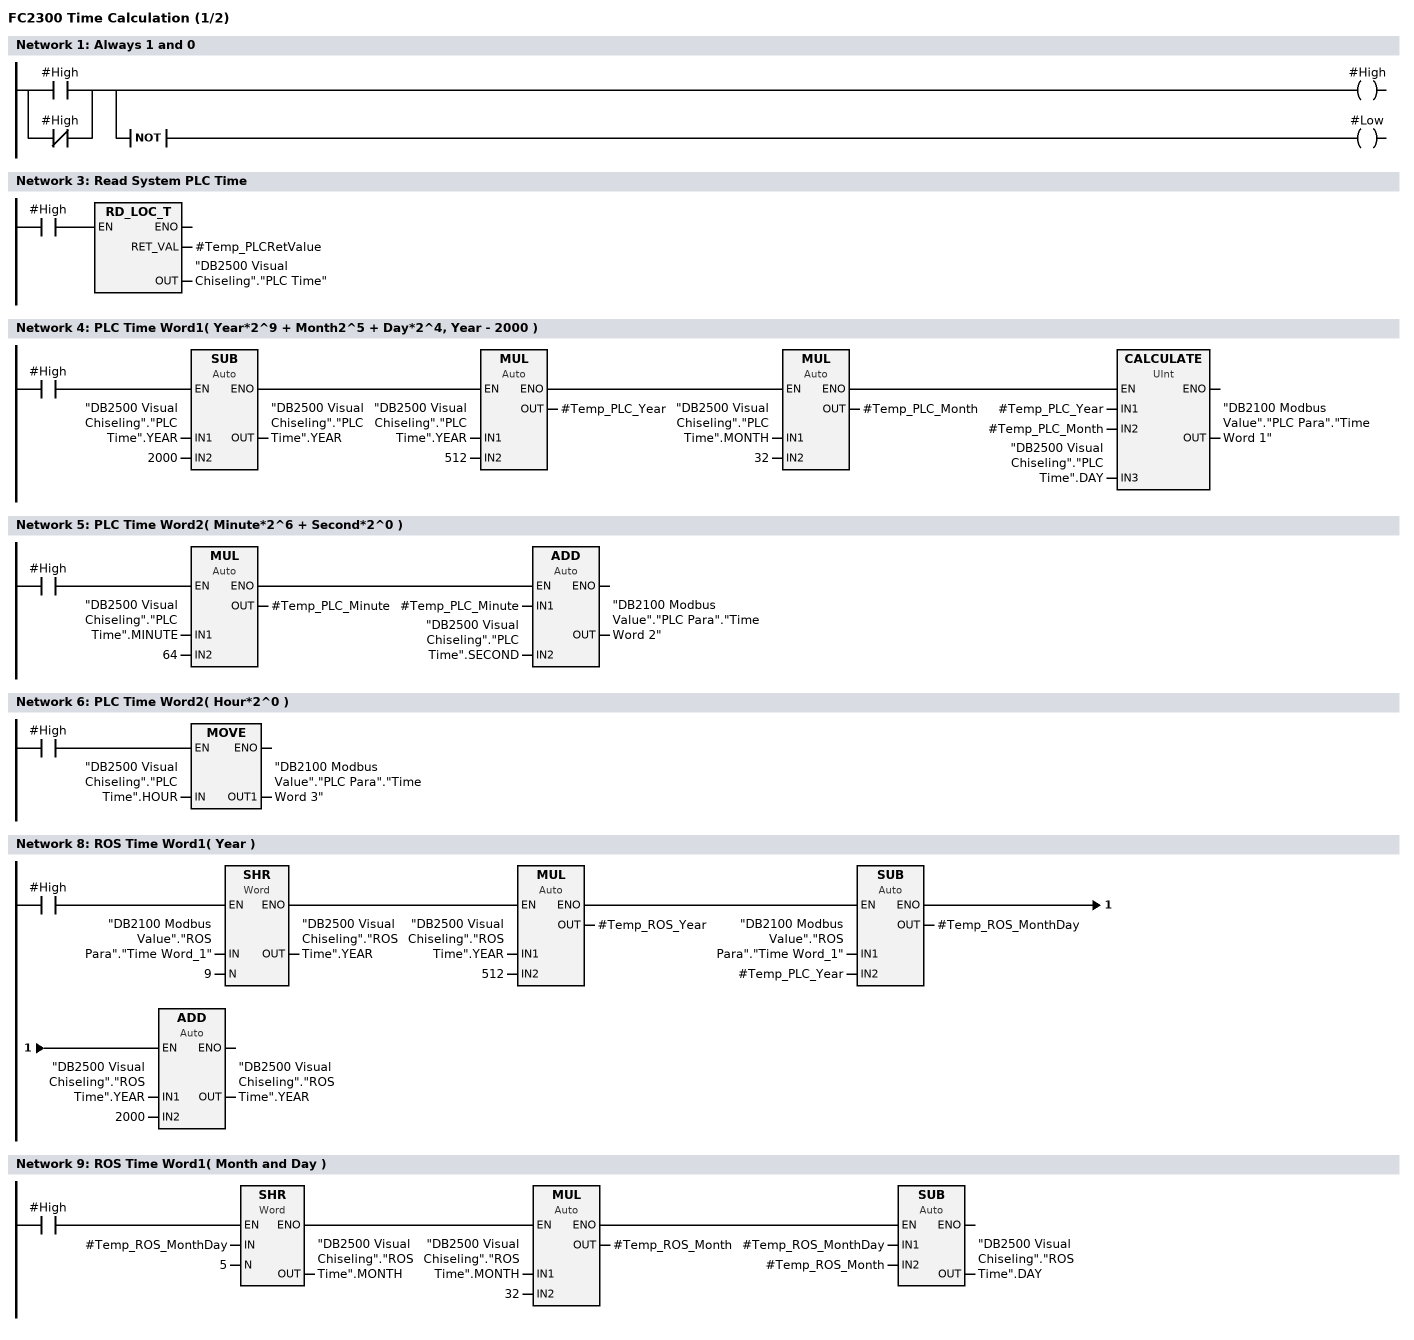
   RUNG wire#powerrail
      Contact( #High )
      wire#w1
      Coil( #High )
   END_RUNG
   RUNG wire#powerrail
      I_Contact( #High )
   END_RUNG wire#w1
   RUNG wire#w1
      Not()
      Coil( #Low )
   END_RUNG
   // the same network as SCL:
   #High := #High OR NOT #High;
   #Low := NOT #High;
END_REGION

REGION Network 2: ############### Write PLC Time To ROS ###############
END_REGION

REGION Network 3: Read System PLC Time
   IF #High THEN #Temp_PLCRetValue := RD_LOC_T(OUT => "DB2500 Visual Chiseling"."PLC Time"); END_IF;
END_REGION

REGION Network 4: PLC Time Word1( Year*2^9 + Month2^5 + Day*2^4, Year - 2000 )
   RUNG wire#powerrail
      Contact( #High )
      Sub(in1 := "DB2500 Visual Chiseling"."PLC Time".YEAR, in2 := 2000, out => "DB2500 Visual Chiseling"."PLC Time".YEAR)
      Mul(in1 := "DB2500 Visual Chiseling"."PLC Time".YEAR, in2 := 512, out => #Temp_PLC_Year)
      Mul(in1 := "DB2500 Visual Chiseling"."PLC Time".MONTH, in2 := 32, out => #Temp_PLC_Month)
      { S7_Templates := "SrcType := UInt"; S7_Expression := "IN1+IN2+IN3" } Calculate(in1 := #Temp_PLC_Year, in2 := #Temp_PLC_Month, in3 := "DB2500 Visual Chiseling"."PLC Time".DAY, out => "DB2100 Modbus Value"."PLC Para"."Time Word 1")
   END_RUNG
   // the same network as SCL:
   IF #High THEN
       "DB2500 Visual Chiseling"."PLC Time".YEAR := "DB2500 Visual Chiseling"."PLC Time".YEAR - 2000;
       #Temp_PLC_Year := "DB2500 Visual Chiseling"."PLC Time".YEAR * 512;
       #Temp_PLC_Month := "DB2500 Visual Chiseling"."PLC Time".MONTH * 32;
       "DB2100 Modbus Value"."PLC Para"."Time Word 1" := #Temp_PLC_Year+#Temp_PLC_Month+"DB2500 Visual Chiseling"."PLC Time".DAY;
   END_IF;
END_REGION

REGION Network 5: PLC Time Word2( Minute*2^6 + Second*2^0 )
   RUNG wire#powerrail
      Contact( #High )
      Mul(in1 := "DB2500 Visual Chiseling"."PLC Time".MINUTE, in2 := 64, out => #Temp_PLC_Minute)
      Add(in1 := #Temp_PLC_Minute, in2 := "DB2500 Visual Chiseling"."PLC Time".SECOND, out => "DB2100 Modbus Value"."PLC Para"."Time Word 2")
   END_RUNG
   // the same network as SCL:
   IF #High THEN
       #Temp_PLC_Minute := "DB2500 Visual Chiseling"."PLC Time".MINUTE * 64;
       "DB2100 Modbus Value"."PLC Para"."Time Word 2" := #Temp_PLC_Minute + "DB2500 Visual Chiseling"."PLC Time".SECOND;
   END_IF;
END_REGION

REGION Network 6: PLC Time Word2( Hour*2^0 )
   RUNG wire#powerrail
      Contact( #High )
      Move(in := "DB2500 Visual Chiseling"."PLC Time".HOUR, out1 => "DB2100 Modbus Value"."PLC Para"."Time Word 3")
   END_RUNG
   // the same network as SCL:
   IF #High THEN
       "DB2100 Modbus Value"."PLC Para"."Time Word 3" := "DB2500 Visual Chiseling"."PLC Time".HOUR;
   END_IF;
END_REGION

REGION Network 7: ############### Read ROS Time To PLC ###############
END_REGION

REGION Network 8: ROS Time Word1( Year )
   RUNG wire#powerrail
      Contact( #High )
      { S7_Templates := "SrcType := Word" } Shr(in := "DB2100 Modbus Value"."ROS Para"."Time Word_1", n := 9, out => "DB2500 Visual Chiseling"."ROS Time".YEAR)
      Mul(in1 := "DB2500 Visual Chiseling"."ROS Time".YEAR, in2 := 512, out => #Temp_ROS_Year)
      Sub(in1 := "DB2100 Modbus Value"."ROS Para"."Time Word_1", in2 := #Temp_PLC_Year, out => #Temp_ROS_MonthDay)
      Add(in1 := "DB2500 Visual Chiseling"."ROS Time".YEAR, in2 := 2000, out => "DB2500 Visual Chiseling"."ROS Time".YEAR)
   END_RUNG
   // the same network as SCL:
   IF #High THEN
       "DB2500 Visual Chiseling"."ROS Time".YEAR := SHR(IN := "DB2100 Modbus Value"."ROS Para"."Time Word_1", N := 9);
       #Temp_ROS_Year := "DB2500 Visual Chiseling"."ROS Time".YEAR * 512;
       #Temp_ROS_MonthDay := "DB2100 Modbus Value"."ROS Para"."Time Word_1" - #Temp_PLC_Year;
       "DB2500 Visual Chiseling"."ROS Time".YEAR := "DB2500 Visual Chiseling"."ROS Time".YEAR + 2000;
   END_IF;
END_REGION

REGION Network 9: ROS Time Word1( Month and Day )
   RUNG wire#powerrail
      Contact( #High )
      { S7_Templates := "SrcType := Word" } Shr(in := #Temp_ROS_MonthDay, n := 5, out => "DB2500 Visual Chiseling"."ROS Time".MONTH)
      Mul(in1 := "DB2500 Visual Chiseling"."ROS Time".MONTH, in2 := 32, out => #Temp_ROS_Month)
      Sub(in1 := #Temp_ROS_MonthDay, in2 := #Temp_ROS_Month, out => "DB2500 Visual Chiseling"."ROS Time".DAY)
   END_RUNG
   // the same network as SCL:
   IF #High THEN
       "DB2500 Visual Chiseling"."ROS Time".MONTH := SHR(IN := #Temp_ROS_MonthDay, N := 5);
       #Temp_ROS_Month := "DB2500 Visual Chiseling"."ROS Time".MONTH * 32;
       "DB2500 Visual Chiseling"."ROS Time".DAY := #Temp_ROS_MonthDay - #Temp_ROS_Month;
   END_IF;
END_REGION

REGION Network 10: ROS Time Word2 ( Minute and Second )
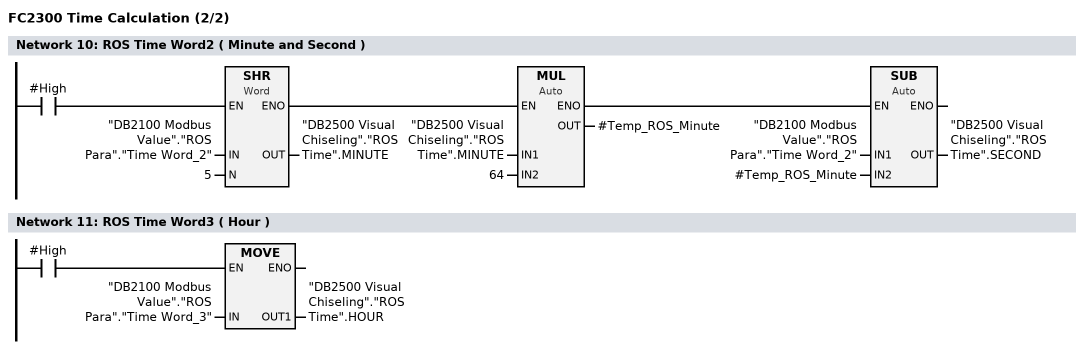
   RUNG wire#powerrail
      Contact( #High )
      { S7_Templates := "SrcType := Word" } Shr(in := "DB2100 Modbus Value"."ROS Para"."Time Word_2", n := 5, out => "DB2500 Visual Chiseling"."ROS Time".MINUTE)
      Mul(in1 := "DB2500 Visual Chiseling"."ROS Time".MINUTE, in2 := 64, out => #Temp_ROS_Minute)
      Sub(in1 := "DB2100 Modbus Value"."ROS Para"."Time Word_2", in2 := #Temp_ROS_Minute, out => "DB2500 Visual Chiseling"."ROS Time".SECOND)
   END_RUNG
   // the same network as SCL:
   IF #High THEN
       "DB2500 Visual Chiseling"."ROS Time".MINUTE := SHR(IN := "DB2100 Modbus Value"."ROS Para"."Time Word_2", N := 5);
       #Temp_ROS_Minute := "DB2500 Visual Chiseling"."ROS Time".MINUTE * 64;
       "DB2500 Visual Chiseling"."ROS Time".SECOND := "DB2100 Modbus Value"."ROS Para"."Time Word_2" - #Temp_ROS_Minute;
   END_IF;
END_REGION

REGION Network 11: ROS Time Word3 ( Hour )
   RUNG wire#powerrail
      Contact( #High )
      Move(in := "DB2100 Modbus Value"."ROS Para"."Time Word_3", out1 => "DB2500 Visual Chiseling"."ROS Time".HOUR)
   END_RUNG
   // the same network as SCL:
   IF #High THEN
       "DB2500 Visual Chiseling"."ROS Time".HOUR := "DB2100 Modbus Value"."ROS Para"."Time Word_3";
   END_IF;
END_REGION

REGION Network 12: ##################### END #####################
END_REGION
END_FUNCTION

FUNCTION "FC2400 Visual Calibration" : Void   // FC2400, LAD
{ S7_Optimized_Access := 'TRUE' }
VERSION : 0.1
   VAR_TEMP
      High : Bool;
      TempPoint_REAL : Struct
         X : Real;
         Y : Real;
         Z : Real;
         "A" : Real;
         "B" : Real;
         C : Real;
      END_STRUCT;
   END_VAR
BEGIN

REGION Network 1: manual into visual calibration mode
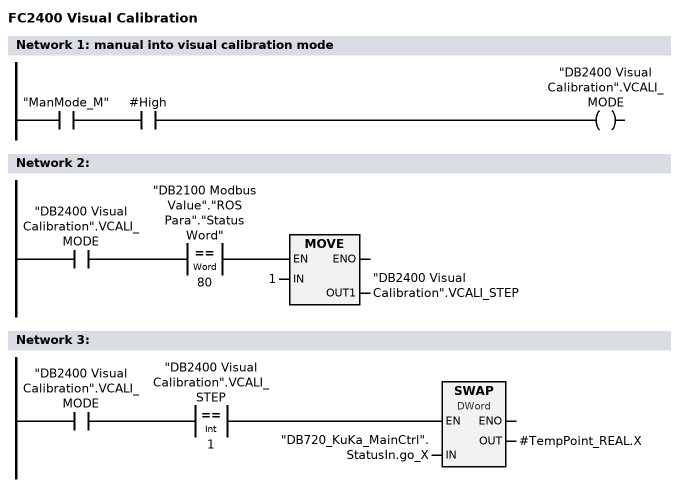
   RUNG wire#powerrail
      Contact( "ManMode_M" )
      Contact( #High )
      Coil( "DB2400 Visual Calibration".VCALI_MODE )
   END_RUNG
   // the same network as SCL:
   "DB2400 Visual Calibration".VCALI_MODE := "ManMode_M" AND #High;
END_REGION

REGION Network 2
   RUNG wire#powerrail
      Contact( "DB2400 Visual Calibration".VCALI_MODE )
      { S7_Templates := "SrcType := Word" } EQ_Contact(in1 := "DB2100 Modbus Value"."ROS Para"."Status Word", in2 := 80)
      Move(in := 1, out1 => "DB2400 Visual Calibration".VCALI_STEP)
   END_RUNG
   // the same network as SCL:
   IF "DB2400 Visual Calibration".VCALI_MODE AND ("DB2100 Modbus Value"."ROS Para"."Status Word" = 80) THEN
       "DB2400 Visual Calibration".VCALI_STEP := 1;
   END_IF;
END_REGION

REGION Network 3
   IF "DB2400 Visual Calibration".VCALI_MODE AND ("DB2400 Visual Calibration".VCALI_STEP = 1) THEN
       #TempPoint_REAL.X := SWAP("DB720_KuKa_MainCtrl".StatusIn.go_X);
   END_IF;
END_REGION
END_FUNCTION

FUNCTION "FC2500 Visual Chiseling" : Void   // FC2500, LAD
TITLE = Program for Visual Gouge
{ S7_Optimized_Access := 'TRUE' }
VERSION : 0.1
// Programmed by Wang Xinyang, 20220610. Any Problem Please Contact Mr.Wang.
   VAR_TEMP
      High : Bool;
      Low : Bool;
      Temp_ResetVChiselRound : Bool;
      Temp_ActivateCam : Bool;
      Temp_ChiselPoint : Int;
      Temp_CamRound : Int;
      RetValue : Array[0..12] of Int;
      Calculation_OffsetMid : Struct
         X0 : DInt;
         X1 : Real;
         Y0 : DInt;
         Y1 : Real;
         Z0 : DInt;
         Z1 : Real;
         A0 : DInt;
         A1 : Real;
         B0 : DInt;
         B1 : Real;
         C0 : DInt;
         C1 : Real;
      END_STRUCT;
      Visual_OffsetMid : Struct
         X0 : DInt;
         X1 : Real;
         Y0 : DInt;
         Y1 : Real;
         Z0 : DInt;
         Z1 : Real;
         A0 : DInt;
         A1 : Real;
         B0 : DInt;
         B1 : Real;
         C0 : DInt;
         C1 : Real;
      END_STRUCT;
   END_VAR
   VAR_TEMP   // added for the SCL form of the ladder/FBD networks
      _w1 : Bool;
      _w2 : Bool;
      _w3 : Bool;
      _w4 : Bool;
      _w5 : Bool;
      _w6 : Bool;
      _w7 : Bool;
   END_VAR
BEGIN

REGION Network 1: Always 1 and 0
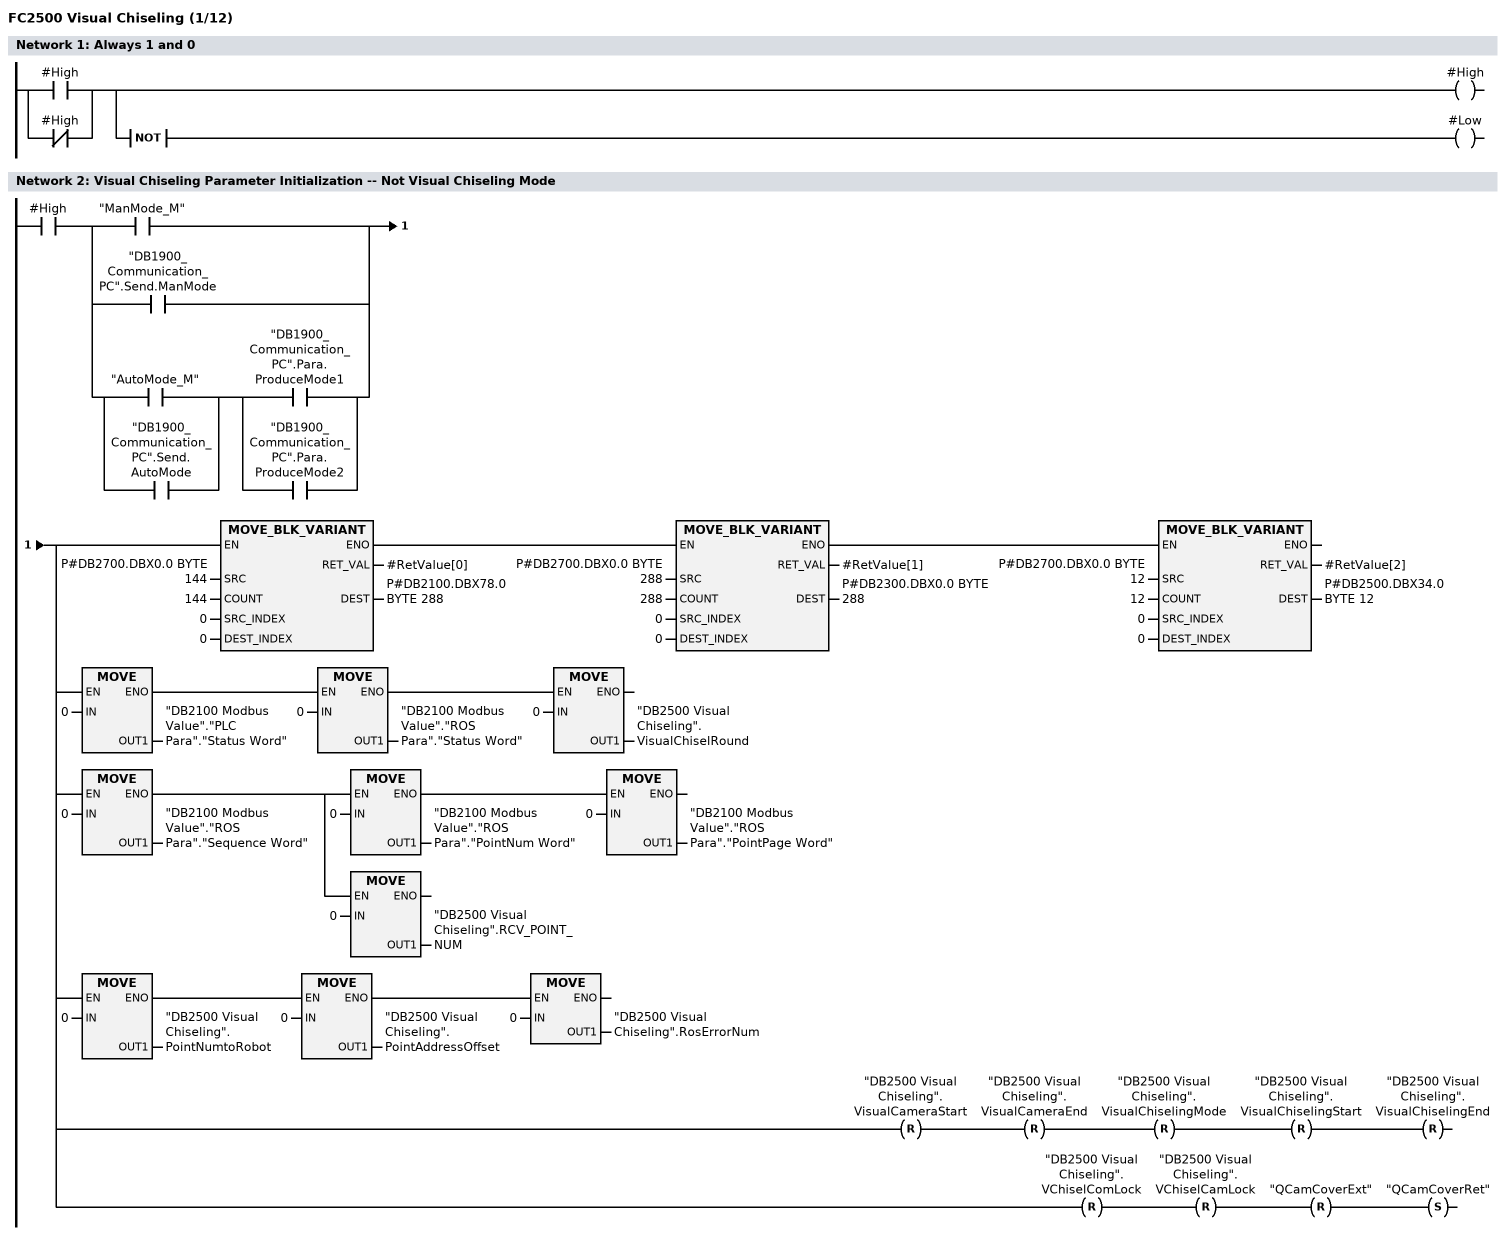
   RUNG wire#powerrail
      Contact( #High )
      wire#w1
      Coil( #High )
   END_RUNG
   RUNG wire#powerrail
      I_Contact( #High )
   END_RUNG wire#w1
   RUNG wire#w1
      Not()
      Coil( #Low )
   END_RUNG
   // the same network as SCL:
   #High := #High OR NOT #High;
   #Low := NOT #High;
END_REGION

REGION Network 2: Visual Chiseling Parameter Initialization -- Not Visual Chiseling Mode
   // ENO of a box is taken as its EN; it also drops when the box reports an error
   #_w1 := #High AND ("ManMode_M" OR "DB1900_Communication_PC".Send.ManMode OR (("AutoMode_M" OR "DB1900_Communication_PC".Send.AutoMode) AND ("DB1900_Communication_PC".Para.ProduceMode1 OR "DB1900_Communication_PC".Para.ProduceMode2)));
   #_w2 := #High AND ("ManMode_M" OR "DB1900_Communication_PC".Send.ManMode OR (("AutoMode_M" OR "DB1900_Communication_PC".Send.AutoMode) AND ("DB1900_Communication_PC".Para.ProduceMode1 OR "DB1900_Communication_PC".Para.ProduceMode2)));
   IF #_w2 THEN
       #RetValue[0] := MOVE_BLK_VARIANT(SRC := P#DB2700.DBX0.0 BYTE 144,
                               COUNT := 144,
                               SRC_INDEX := 0,
                               DEST_INDEX := 0,
                               DEST => P#DB2100.DBX78.0 BYTE 288);
       #RetValue[1] := MOVE_BLK_VARIANT(SRC := P#DB2700.DBX0.0 BYTE 288,
                               COUNT := 288,
                               SRC_INDEX := 0,
                               DEST_INDEX := 0,
                               DEST => P#DB2300.DBX0.0 BYTE 288);
       #RetValue[2] := MOVE_BLK_VARIANT(SRC := P#DB2700.DBX0.0 BYTE 12,
                               COUNT := 12,
                               SRC_INDEX := 0,
                               DEST_INDEX := 0,
                               DEST => P#DB2500.DBX34.0 BYTE 12);
   END_IF;
   IF #_w1 THEN
       "DB2100 Modbus Value"."PLC Para"."Status Word" := 0;
       "DB2100 Modbus Value"."ROS Para"."Status Word" := 0;
       "DB2500 Visual Chiseling".VisualChiselRound := 0;
       "DB2100 Modbus Value"."ROS Para"."Sequence Word" := 0;
       "DB2100 Modbus Value"."ROS Para"."PointNum Word" := 0;
       "DB2100 Modbus Value"."ROS Para"."PointPage Word" := 0;
       "DB2500 Visual Chiseling".RCV_POINT_NUM := 0;
       "DB2500 Visual Chiseling".PointNumtoRobot := 0;
       "DB2500 Visual Chiseling".PointAddressOffset := 0;
       "DB2500 Visual Chiseling".RosErrorNum := 0;
       "DB2500 Visual Chiseling".VisualCameraStart := FALSE;
       "DB2500 Visual Chiseling".VisualCameraEnd := FALSE;
       "DB2500 Visual Chiseling".VisualChiselingMode := FALSE;
       "DB2500 Visual Chiseling".VisualChiselingStart := FALSE;
       "DB2500 Visual Chiseling".VisualChiselingEnd := FALSE;
       "DB2500 Visual Chiseling".VChiselComLock := FALSE;
       "DB2500 Visual Chiseling".VChiselCamLock := FALSE;
       "QCamCoverExt" := FALSE;
       "QCamCoverRet" := TRUE;
   END_IF;
END_REGION

REGION Network 3: ############### Auto Visual Camera Function ###############
END_REGION

REGION Network 4: Step0: Activate Visual Chiseling Mode
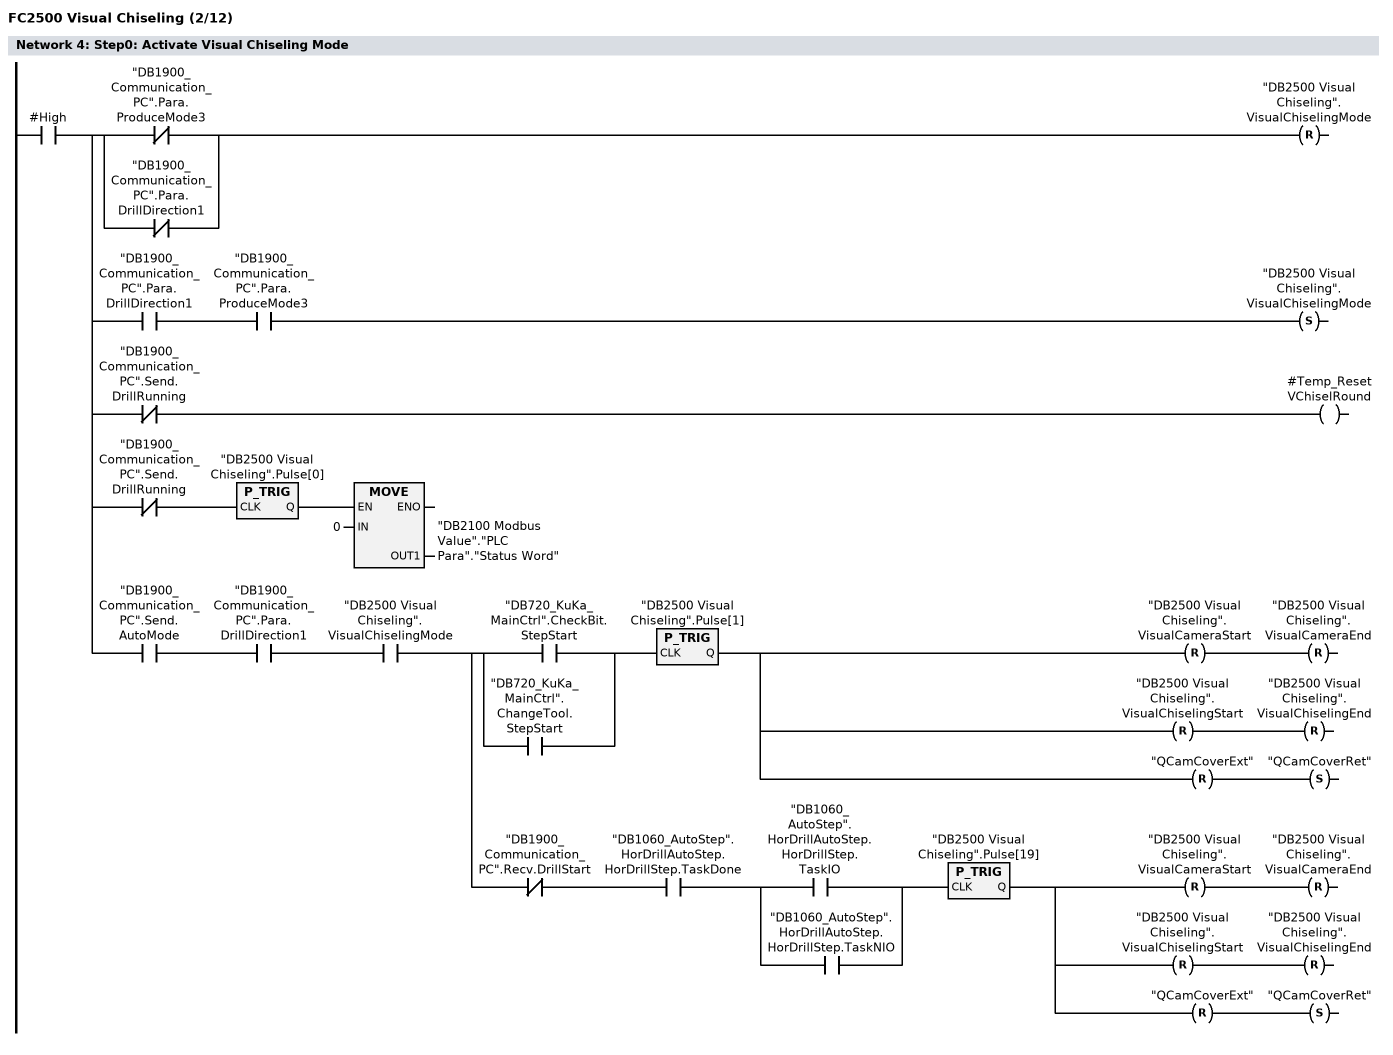
   RUNG wire#powerrail
      Contact( #High )
      wire#w1
      I_Contact( "DB1900_Communication_PC".Para.ProduceMode3 )
      wire#w2
      R_Coil( "DB2500 Visual Chiseling".VisualChiselingMode )
   END_RUNG
   RUNG wire#w1
      I_Contact( "DB1900_Communication_PC".Para.DrillDirection1 )
   END_RUNG wire#w2
   RUNG wire#w1
      Contact( "DB1900_Communication_PC".Para.DrillDirection1 )
      Contact( "DB1900_Communication_PC".Para.ProduceMode3 )
      S_Coil( "DB2500 Visual Chiseling".VisualChiselingMode )
   END_RUNG
   RUNG wire#w1
      I_Contact( "DB1900_Communication_PC".Send.DrillRunning )
      Coil( #Temp_ResetVChiselRound )
   END_RUNG
   RUNG wire#w1
      I_Contact( "DB1900_Communication_PC".Send.DrillRunning )
      P_Trig( "DB2500 Visual Chiseling".Pulse[0] )
      Move(in := 0, out1 => "DB2100 Modbus Value"."PLC Para"."Status Word")
   END_RUNG
   RUNG wire#w1
      Contact( "DB1900_Communication_PC".Send.AutoMode )
      Contact( "DB1900_Communication_PC".Para.DrillDirection1 )
      Contact( "DB2500 Visual Chiseling".VisualChiselingMode )
      wire#w3
      Contact( "DB720_KuKa_MainCtrl".CheckBit.StepStart )
      wire#w4
      P_Trig( "DB2500 Visual Chiseling".Pulse[1] )
      wire#w5
      R_Coil( "DB2500 Visual Chiseling".VisualCameraStart )
      R_Coil( "DB2500 Visual Chiseling".VisualCameraEnd )
   END_RUNG
   RUNG wire#w3
      Contact( "DB720_KuKa_MainCtrl".ChangeTool.StepStart )
   END_RUNG wire#w4
   RUNG wire#w5
      R_Coil( "DB2500 Visual Chiseling".VisualChiselingStart )
      R_Coil( "DB2500 Visual Chiseling".VisualChiselingEnd )
   END_RUNG
   RUNG wire#w5
      R_Coil( "QCamCoverExt" )
      S_Coil( "QCamCoverRet" )
   END_RUNG
   RUNG wire#w3
      I_Contact( "DB1900_Communication_PC".Recv.DrillStart )
      Contact( "DB1060_AutoStep".HorDrillAutoStep.HorDrillStep.TaskDone )
      wire#w6
      Contact( "DB1060_AutoStep".HorDrillAutoStep.HorDrillStep.TaskIO )
      wire#w7
      P_Trig( "DB2500 Visual Chiseling".Pulse[19] )
      wire#w8
      R_Coil( "DB2500 Visual Chiseling".VisualCameraStart )
      R_Coil( "DB2500 Visual Chiseling".VisualCameraEnd )
   END_RUNG
   RUNG wire#w6
      Contact( "DB1060_AutoStep".HorDrillAutoStep.HorDrillStep.TaskNIO )
   END_RUNG wire#w7
   RUNG wire#w8
      R_Coil( "DB2500 Visual Chiseling".VisualChiselingStart )
      R_Coil( "DB2500 Visual Chiseling".VisualChiselingEnd )
   END_RUNG
   RUNG wire#w8
      R_Coil( "QCamCoverExt" )
      S_Coil( "QCamCoverRet" )
   END_RUNG
   // the same network as SCL:
   IF #High AND (NOT "DB1900_Communication_PC".Para.ProduceMode3 OR NOT "DB1900_Communication_PC".Para.DrillDirection1) THEN
       "DB2500 Visual Chiseling".VisualChiselingMode := FALSE;
   END_IF;
   IF #High AND "DB1900_Communication_PC".Para.DrillDirection1 AND "DB1900_Communication_PC".Para.ProduceMode3 THEN
       "DB2500 Visual Chiseling".VisualChiselingMode := TRUE;
   END_IF;
   #Temp_ResetVChiselRound := #High AND NOT "DB1900_Communication_PC".Send.DrillRunning;
   #_w1 := #High AND NOT "DB1900_Communication_PC".Send.DrillRunning;
   #_w2 := #_w1 AND NOT "DB2500 Visual Chiseling".Pulse[0];   // rising edge
   "DB2500 Visual Chiseling".Pulse[0] := #_w1;
   IF #_w2 THEN "DB2100 Modbus Value"."PLC Para"."Status Word" := 0; END_IF;
   #_w3 := #High AND "DB1900_Communication_PC".Send.AutoMode AND "DB1900_Communication_PC".Para.DrillDirection1 AND "DB2500 Visual Chiseling".VisualChiselingMode;
   #_w4 := #_w3 AND ("DB720_KuKa_MainCtrl".CheckBit.StepStart OR "DB720_KuKa_MainCtrl".ChangeTool.StepStart);
   #_w5 := #_w4 AND NOT "DB2500 Visual Chiseling".Pulse[1];   // rising edge
   "DB2500 Visual Chiseling".Pulse[1] := #_w4;
   IF #_w5 THEN
       "DB2500 Visual Chiseling".VisualCameraStart := FALSE;
       "DB2500 Visual Chiseling".VisualCameraEnd := FALSE;
       "DB2500 Visual Chiseling".VisualChiselingStart := FALSE;
       "DB2500 Visual Chiseling".VisualChiselingEnd := FALSE;
       "QCamCoverExt" := FALSE;
       "QCamCoverRet" := TRUE;
   END_IF;
   #_w6 := #_w3 AND NOT "DB1900_Communication_PC".Recv.DrillStart AND "DB1060_AutoStep".HorDrillAutoStep.HorDrillStep.TaskDone AND ("DB1060_AutoStep".HorDrillAutoStep.HorDrillStep.TaskIO OR "DB1060_AutoStep".HorDrillAutoStep.HorDrillStep.TaskNIO);
   #_w7 := #_w6 AND NOT "DB2500 Visual Chiseling".Pulse[19];   // rising edge
   "DB2500 Visual Chiseling".Pulse[19] := #_w6;
   IF #_w7 THEN
       "DB2500 Visual Chiseling".VisualCameraStart := FALSE;
       "DB2500 Visual Chiseling".VisualCameraEnd := FALSE;
       "DB2500 Visual Chiseling".VisualChiselingStart := FALSE;
       "DB2500 Visual Chiseling".VisualChiselingEnd := FALSE;
       "QCamCoverExt" := FALSE;
       "QCamCoverRet" := TRUE;
   END_IF;
END_REGION

REGION Network 5: Step0: Auto Visual Chiseling Function Start
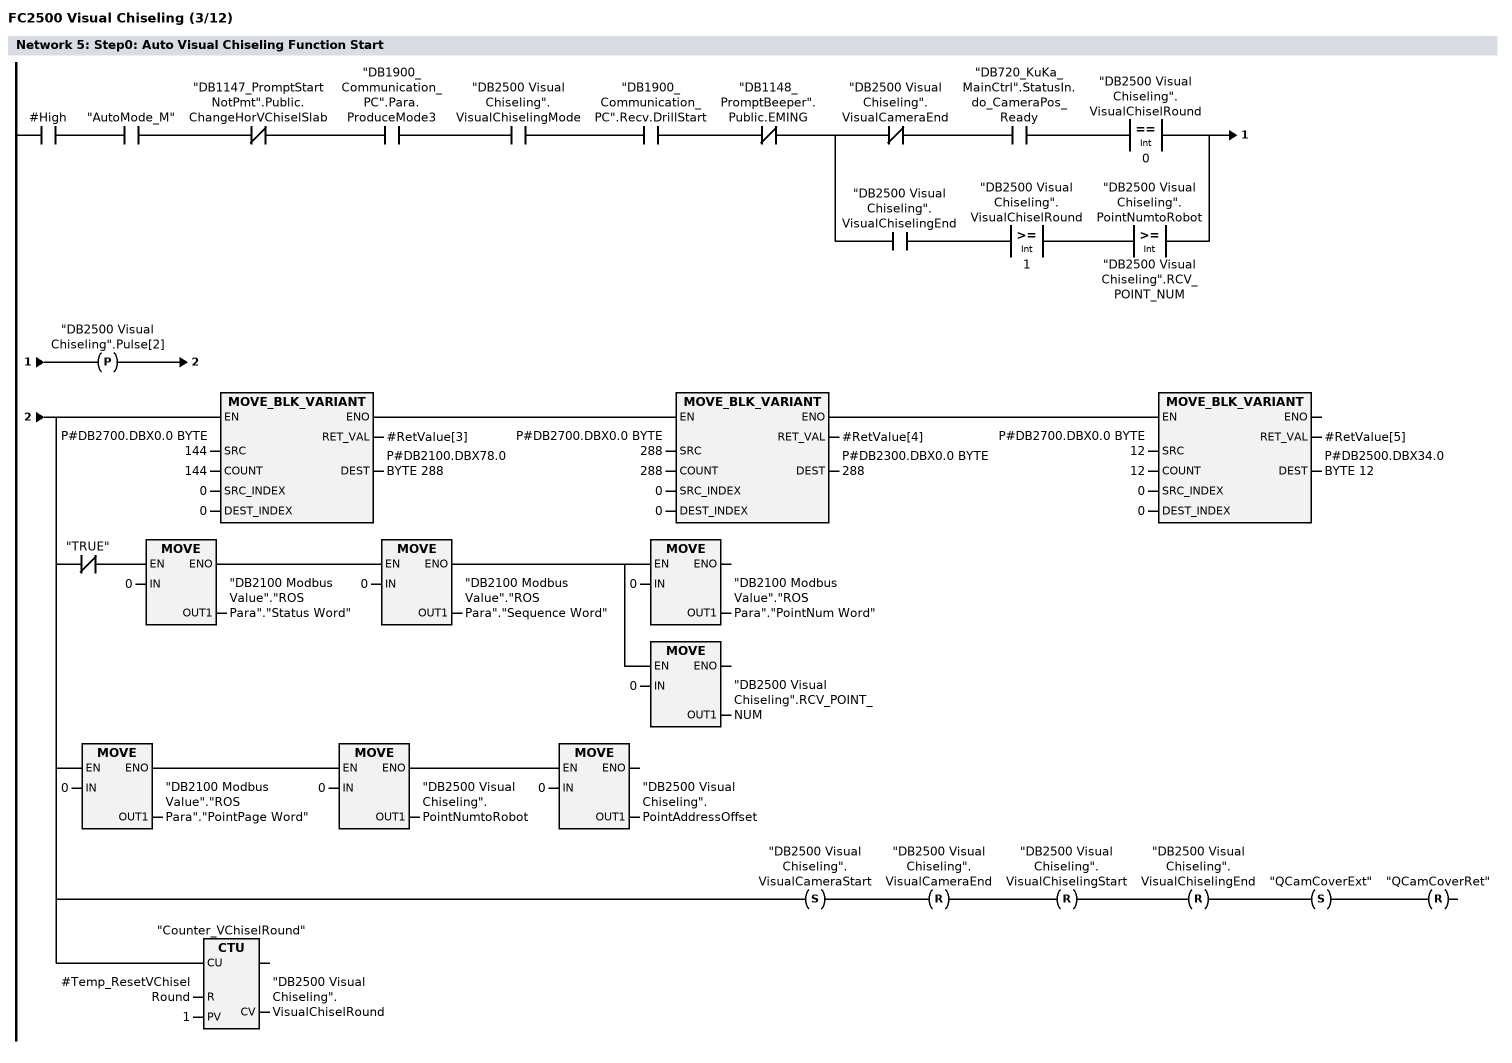
   // ENO of a box is taken as its EN; it also drops when the box reports an error
   #_w1 := #High AND "AutoMode_M" AND NOT "DB1147_PromptStartNotPmt".Public.ChangeHorVChiselSlab AND "DB1900_Communication_PC".Para.ProduceMode3 AND "DB2500 Visual Chiseling".VisualChiselingMode AND "DB1900_Communication_PC".Recv.DrillStart AND NOT "DB1148_PromptBeeper".Public.EMING AND ((NOT "DB2500 Visual Chiseling".VisualCameraEnd AND "DB720_KuKa_MainCtrl".StatusIn.do_CameraPos_Ready AND ("DB2500 Visual Chiseling".VisualChiselRound = 0)) OR ("DB2500 Visual Chiseling".VisualChiselingEnd AND ("DB2500 Visual Chiseling".VisualChiselRound >= 1) AND ("DB2500 Visual Chiseling".PointNumtoRobot >= "DB2500 Visual Chiseling".RCV_POINT_NUM)));
   #_w2 := #_w1 AND NOT "DB2500 Visual Chiseling".Pulse[2];   // rising edge
   "DB2500 Visual Chiseling".Pulse[2] := #_w1;
   IF #_w2 THEN
       #RetValue[3] := MOVE_BLK_VARIANT(SRC := P#DB2700.DBX0.0 BYTE 144,
                               COUNT := 144,
                               SRC_INDEX := 0,
                               DEST_INDEX := 0,
                               DEST => P#DB2100.DBX78.0 BYTE 288);
       #RetValue[4] := MOVE_BLK_VARIANT(SRC := P#DB2700.DBX0.0 BYTE 288,
                               COUNT := 288,
                               SRC_INDEX := 0,
                               DEST_INDEX := 0,
                               DEST => P#DB2300.DBX0.0 BYTE 288);
       #RetValue[5] := MOVE_BLK_VARIANT(SRC := P#DB2700.DBX0.0 BYTE 12,
                               COUNT := 12,
                               SRC_INDEX := 0,
                               DEST_INDEX := 0,
                               DEST => P#DB2500.DBX34.0 BYTE 12);
   END_IF;
   IF #_w2 AND NOT "TRUE" THEN
       "DB2100 Modbus Value"."ROS Para"."Status Word" := 0;
       "DB2100 Modbus Value"."ROS Para"."Sequence Word" := 0;
       "DB2100 Modbus Value"."ROS Para"."PointNum Word" := 0;
       "DB2500 Visual Chiseling".RCV_POINT_NUM := 0;
   END_IF;
   IF #_w2 THEN
       "DB2100 Modbus Value"."ROS Para"."PointPage Word" := 0;
       "DB2500 Visual Chiseling".PointNumtoRobot := 0;
       "DB2500 Visual Chiseling".PointAddressOffset := 0;
       "DB2500 Visual Chiseling".VisualCameraStart := TRUE;
       "DB2500 Visual Chiseling".VisualCameraEnd := FALSE;
       "DB2500 Visual Chiseling".VisualChiselingStart := FALSE;
       "DB2500 Visual Chiseling".VisualChiselingEnd := FALSE;
       "QCamCoverExt" := TRUE;
       "QCamCoverRet" := FALSE;
   END_IF;
   "Counter_VChiselRound".CTU(CU := #_w2,
                           R := #Temp_ResetVChiselRound,
                           PV := 1,
                           CV => "DB2500 Visual Chiseling".VisualChiselRound);
END_REGION

REGION Network 6: Step2: Request Activate Camera | PLC Status Word:100
   // StatusWord 100 : Activate Camera in Transition Position,
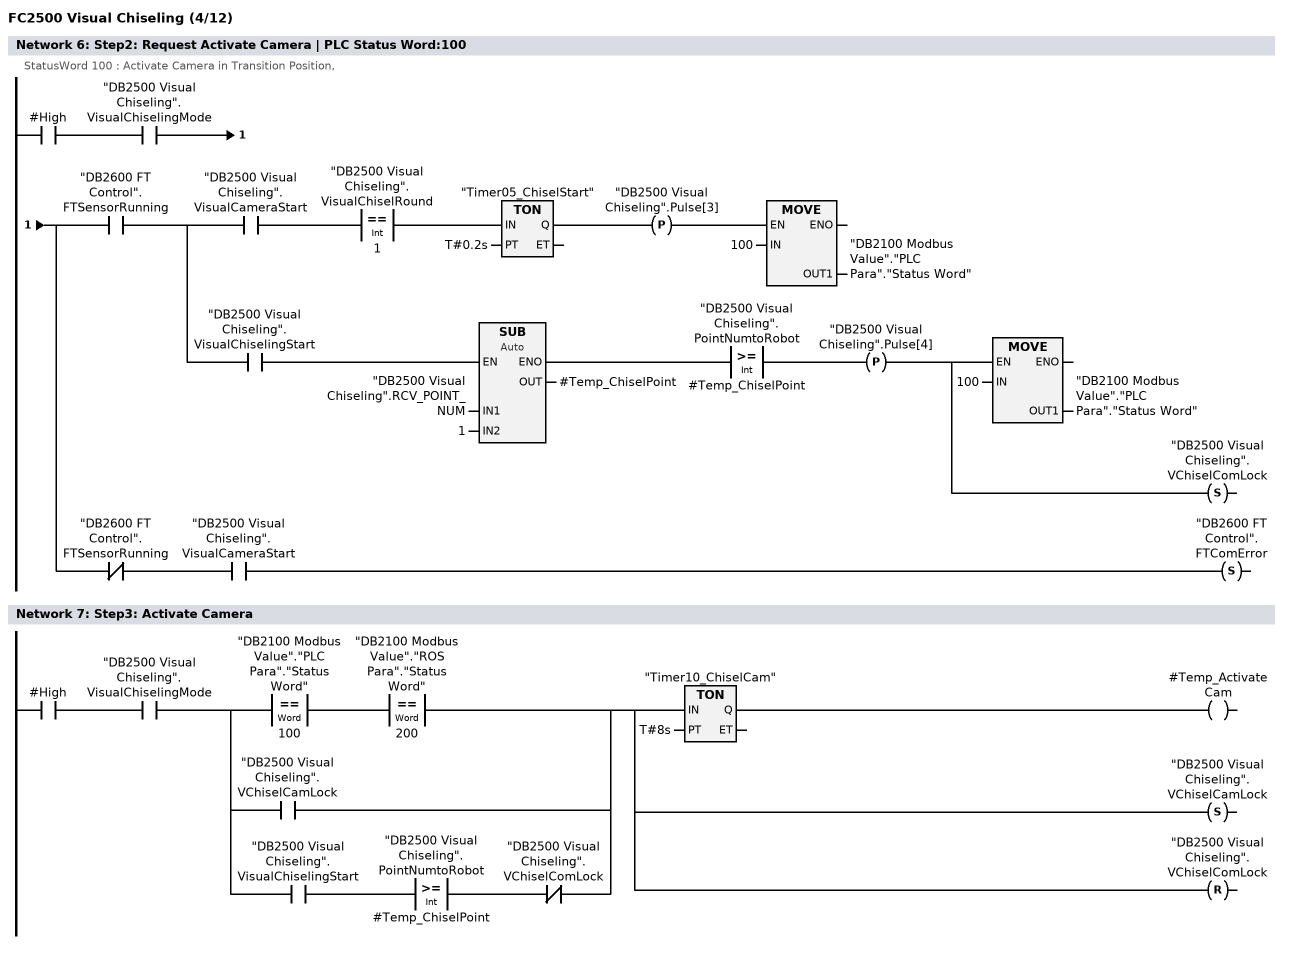
   #_w1 := #High AND "DB2500 Visual Chiseling".VisualChiselingMode;
   #_w2 := #_w1 AND "DB2600 FT Control".FTSensorRunning;
   "Timer05_ChiselStart".TON(IN := #_w2 AND "DB2500 Visual Chiseling".VisualCameraStart AND ("DB2500 Visual Chiseling".VisualChiselRound = 1),
                           PT := T#0.2s);
   #_w3 := "Timer05_ChiselStart".Q AND NOT "DB2500 Visual Chiseling".Pulse[3];   // rising edge
   "DB2500 Visual Chiseling".Pulse[3] := "Timer05_ChiselStart".Q;
   IF #_w3 THEN "DB2100 Modbus Value"."PLC Para"."Status Word" := 100; END_IF;
   #_w4 := #_w2 AND "DB2500 Visual Chiseling".VisualChiselingStart;
   IF #_w4 THEN #Temp_ChiselPoint := "DB2500 Visual Chiseling".RCV_POINT_NUM - 1; END_IF;
   #_w5 := #_w4 AND ("DB2500 Visual Chiseling".PointNumtoRobot >= #Temp_ChiselPoint);
   #_w6 := #_w5 AND NOT "DB2500 Visual Chiseling".Pulse[4];   // rising edge
   "DB2500 Visual Chiseling".Pulse[4] := #_w5;
   IF #_w6 THEN
       "DB2100 Modbus Value"."PLC Para"."Status Word" := 100;
       "DB2500 Visual Chiseling".VChiselComLock := TRUE;
   END_IF;
   IF #_w1 AND NOT "DB2600 FT Control".FTSensorRunning AND "DB2500 Visual Chiseling".VisualCameraStart THEN
       "DB2600 FT Control".FTComError := TRUE;
   END_IF;
END_REGION

REGION Network 7: Step3: Activate Camera
   #_w1 := #High AND "DB2500 Visual Chiseling".VisualChiselingMode AND ((("DB2100 Modbus Value"."PLC Para"."Status Word" = 100) AND ("DB2100 Modbus Value"."ROS Para"."Status Word" = 200)) OR "DB2500 Visual Chiseling".VChiselCamLock OR ("DB2500 Visual Chiseling".VisualChiselingStart AND ("DB2500 Visual Chiseling".PointNumtoRobot >= #Temp_ChiselPoint) AND NOT "DB2500 Visual Chiseling".VChiselComLock));
   "Timer10_ChiselCam".TON(IN := #_w1, PT := T#8s);
   #Temp_ActivateCam := "Timer10_ChiselCam".Q;
   IF #_w1 THEN
       "DB2500 Visual Chiseling".VChiselCamLock := TRUE;
       "DB2500 Visual Chiseling".VChiselComLock := FALSE;
   END_IF;
END_REGION

REGION Network 8: Step3: Request ROS Take Photos and Calculate Point Data | PLC Status Word:110 ROS Status Word: 200
   // StatusWord110:  Request ROS Take Photos When Camera is Ready.
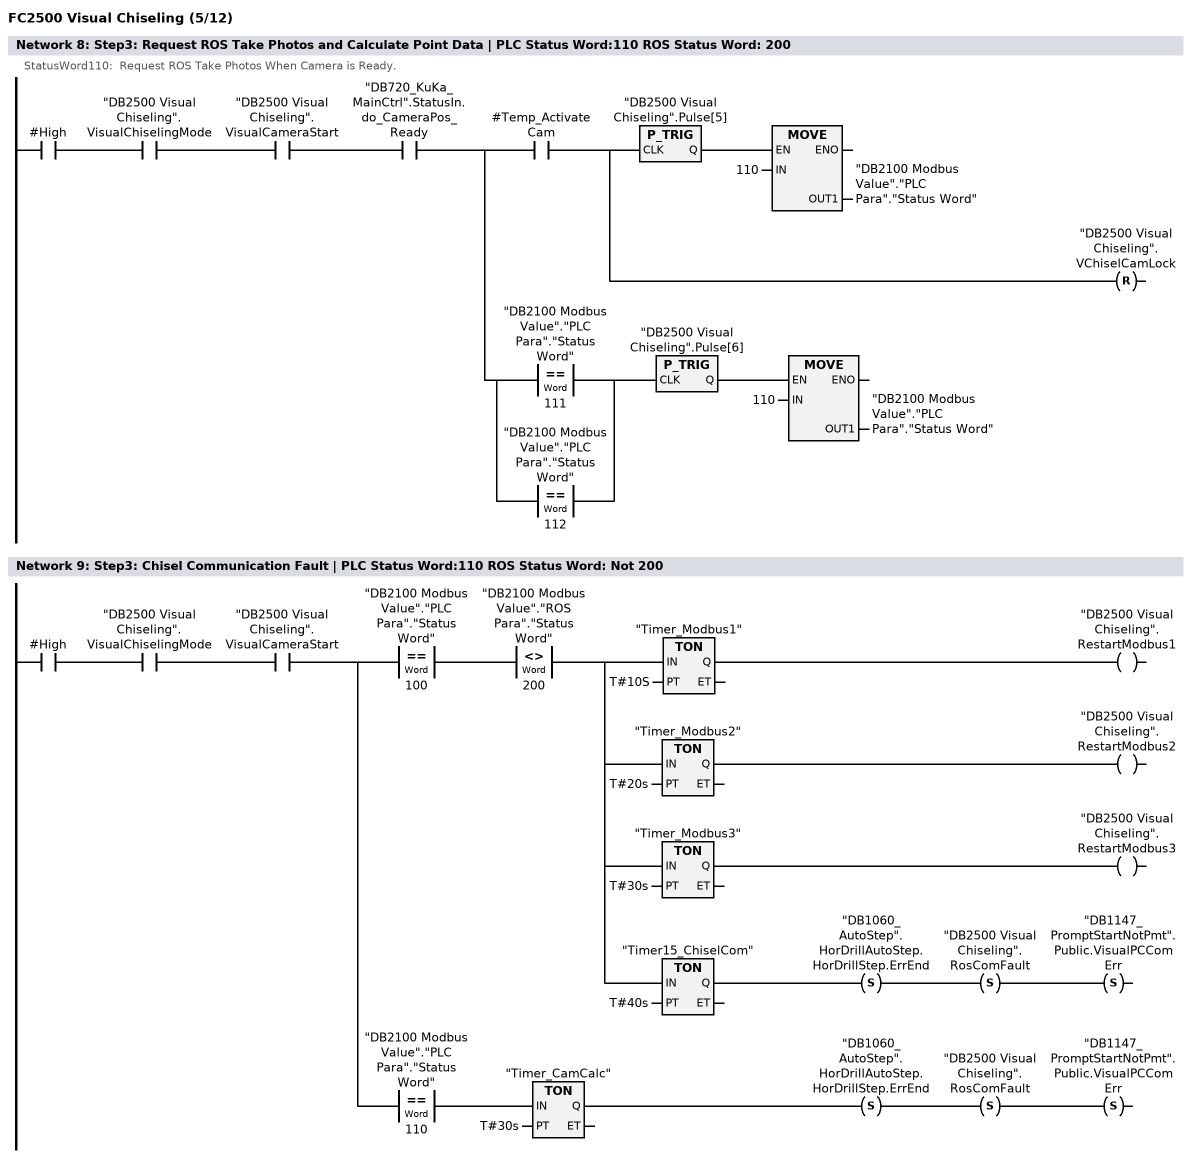
   RUNG wire#powerrail
      Contact( #High )
      Contact( "DB2500 Visual Chiseling".VisualChiselingMode )
      Contact( "DB2500 Visual Chiseling".VisualCameraStart )
      Contact( "DB720_KuKa_MainCtrl".StatusIn.do_CameraPos_Ready )
      wire#w1
      Contact( #Temp_ActivateCam )
      wire#w2
      P_Trig( "DB2500 Visual Chiseling".Pulse[5] )
      Move(in := 110, out1 => "DB2100 Modbus Value"."PLC Para"."Status Word")
   END_RUNG
   RUNG wire#w2
      R_Coil( "DB2500 Visual Chiseling".VChiselCamLock )
   END_RUNG
   RUNG wire#w1
      { S7_Templates := "SrcType := Word" } EQ_Contact(in1 := "DB2100 Modbus Value"."PLC Para"."Status Word", in2 := 111)
      wire#w3
      P_Trig( "DB2500 Visual Chiseling".Pulse[6] )
      Move(in := 110, out1 => "DB2100 Modbus Value"."PLC Para"."Status Word")
   END_RUNG
   RUNG wire#w1
      { S7_Templates := "SrcType := Word" } EQ_Contact(in1 := "DB2100 Modbus Value"."PLC Para"."Status Word", in2 := 112)
   END_RUNG wire#w3
   // the same network as SCL:
   #_w1 := #High AND "DB2500 Visual Chiseling".VisualChiselingMode AND "DB2500 Visual Chiseling".VisualCameraStart AND "DB720_KuKa_MainCtrl".StatusIn.do_CameraPos_Ready;
   #_w2 := #_w1 AND #Temp_ActivateCam;
   #_w3 := #_w2 AND NOT "DB2500 Visual Chiseling".Pulse[5];   // rising edge
   "DB2500 Visual Chiseling".Pulse[5] := #_w2;
   IF #_w3 THEN "DB2100 Modbus Value"."PLC Para"."Status Word" := 110; END_IF;
   IF #_w2 THEN "DB2500 Visual Chiseling".VChiselCamLock := FALSE; END_IF;
   #_w4 := #_w1 AND (("DB2100 Modbus Value"."PLC Para"."Status Word" = 111) OR ("DB2100 Modbus Value"."PLC Para"."Status Word" = 112));
   #_w5 := #_w4 AND NOT "DB2500 Visual Chiseling".Pulse[6];   // rising edge
   "DB2500 Visual Chiseling".Pulse[6] := #_w4;
   IF #_w5 THEN "DB2100 Modbus Value"."PLC Para"."Status Word" := 110; END_IF;
END_REGION

REGION Network 9: Step3: Chisel Communication Fault | PLC Status Word:110 ROS Status Word: Not 200
   #_w1 := #High AND "DB2500 Visual Chiseling".VisualChiselingMode AND "DB2500 Visual Chiseling".VisualCameraStart;
   #_w2 := #_w1 AND ("DB2100 Modbus Value"."PLC Para"."Status Word" = 100) AND ("DB2100 Modbus Value"."ROS Para"."Status Word" <> 200);
   "Timer_Modbus1".TON(IN := #_w2, PT := T#10S);
   "DB2500 Visual Chiseling".RestartModbus1 := "Timer_Modbus1".Q;
   "Timer_Modbus2".TON(IN := #_w2, PT := T#20s);
   "DB2500 Visual Chiseling".RestartModbus2 := "Timer_Modbus2".Q;
   "Timer_Modbus3".TON(IN := #_w2, PT := T#30s);
   "DB2500 Visual Chiseling".RestartModbus3 := "Timer_Modbus3".Q;
   "Timer15_ChiselCom".TON(IN := #_w2, PT := T#40s);
   IF "Timer15_ChiselCom".Q THEN
       "DB1060_AutoStep".HorDrillAutoStep.HorDrillStep.ErrEnd := TRUE;
       "DB2500 Visual Chiseling".RosComFault := TRUE;
       "DB1147_PromptStartNotPmt".Public.VisualPCComErr := TRUE;
   END_IF;
   "Timer_CamCalc".TON(IN := #_w1 AND ("DB2100 Modbus Value"."PLC Para"."Status Word" = 110), PT := T#30s);
   IF "Timer_CamCalc".Q THEN
       "DB1060_AutoStep".HorDrillAutoStep.HorDrillStep.ErrEnd := TRUE;
       "DB2500 Visual Chiseling".RosComFault := TRUE;
       "DB1147_PromptStartNotPmt".Public.VisualPCComErr := TRUE;
   END_IF;
END_REGION

REGION Network 10: Step5: Read Page1 Point Data From ROS, Save to DB2300 | PLC Status Word:110 ROS Status Word: 210
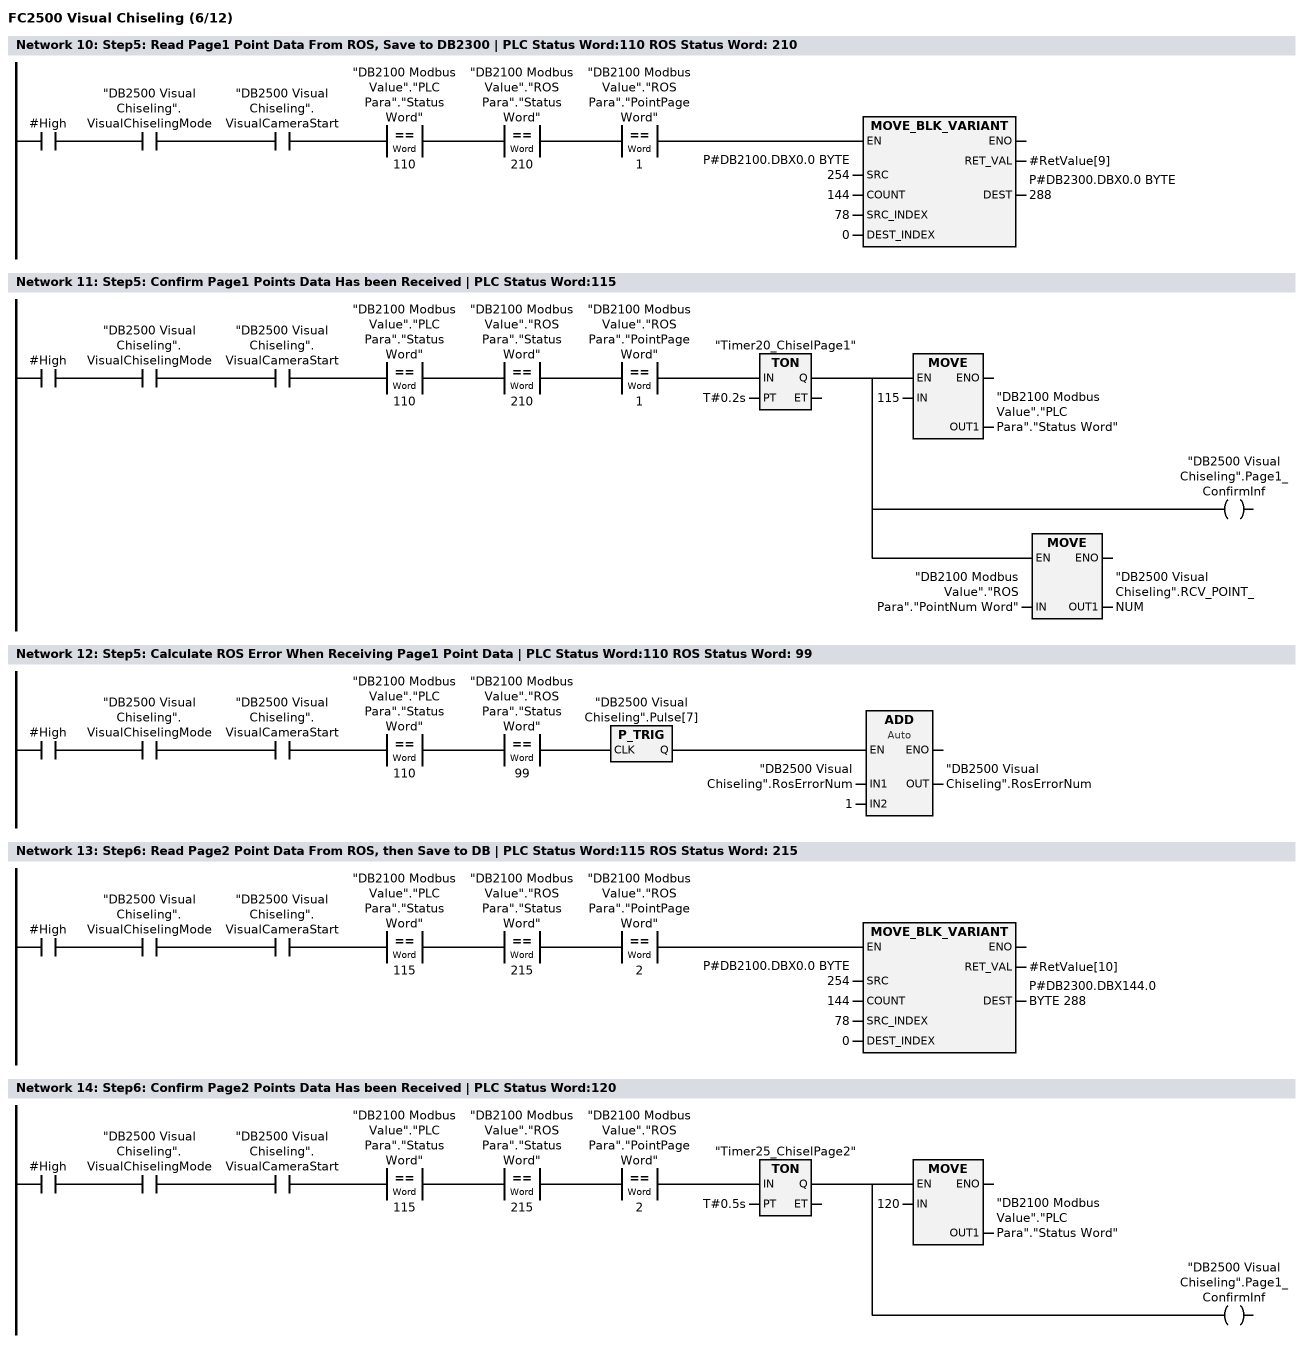
   IF #High AND "DB2500 Visual Chiseling".VisualChiselingMode AND "DB2500 Visual Chiseling".VisualCameraStart AND ("DB2100 Modbus Value"."PLC Para"."Status Word" = 110) AND ("DB2100 Modbus Value"."ROS Para"."Status Word" = 210) AND ("DB2100 Modbus Value"."ROS Para"."PointPage Word" = 1) THEN
       #RetValue[9] := MOVE_BLK_VARIANT(SRC := P#DB2100.DBX0.0 BYTE 254,
                               COUNT := 144,
                               SRC_INDEX := 78,
                               DEST_INDEX := 0,
                               DEST => P#DB2300.DBX0.0 BYTE 288);
   END_IF;
END_REGION

REGION Network 11: Step5: Confirm Page1 Points Data Has been Received | PLC Status Word:115
   "Timer20_ChiselPage1".TON(IN := #High AND "DB2500 Visual Chiseling".VisualChiselingMode AND "DB2500 Visual Chiseling".VisualCameraStart AND ("DB2100 Modbus Value"."PLC Para"."Status Word" = 110) AND ("DB2100 Modbus Value"."ROS Para"."Status Word" = 210) AND ("DB2100 Modbus Value"."ROS Para"."PointPage Word" = 1),
                           PT := T#0.2s);
   IF "Timer20_ChiselPage1".Q THEN "DB2100 Modbus Value"."PLC Para"."Status Word" := 115; END_IF;
   "DB2500 Visual Chiseling".Page1_ConfirmInf := "Timer20_ChiselPage1".Q;
   IF "Timer20_ChiselPage1".Q THEN
       "DB2500 Visual Chiseling".RCV_POINT_NUM := "DB2100 Modbus Value"."ROS Para"."PointNum Word";
   END_IF;
END_REGION

REGION Network 12: Step5: Calculate ROS Error When Receiving Page1 Point Data | PLC Status Word:110 ROS Status Word: 99
   RUNG wire#powerrail
      Contact( #High )
      Contact( "DB2500 Visual Chiseling".VisualChiselingMode )
      Contact( "DB2500 Visual Chiseling".VisualCameraStart )
      { S7_Templates := "SrcType := Word" } EQ_Contact(in1 := "DB2100 Modbus Value"."PLC Para"."Status Word", in2 := 110)
      { S7_Templates := "SrcType := Word" } EQ_Contact(in1 := "DB2100 Modbus Value"."ROS Para"."Status Word", in2 := 99)
      P_Trig( "DB2500 Visual Chiseling".Pulse[7] )
      Add(in1 := "DB2500 Visual Chiseling".RosErrorNum, in2 := 1, out => "DB2500 Visual Chiseling".RosErrorNum)
   END_RUNG
   // the same network as SCL:
   #_w1 := #High AND "DB2500 Visual Chiseling".VisualChiselingMode AND "DB2500 Visual Chiseling".VisualCameraStart AND ("DB2100 Modbus Value"."PLC Para"."Status Word" = 110) AND ("DB2100 Modbus Value"."ROS Para"."Status Word" = 99);
   #_w2 := #_w1 AND NOT "DB2500 Visual Chiseling".Pulse[7];   // rising edge
   "DB2500 Visual Chiseling".Pulse[7] := #_w1;
   IF #_w2 THEN "DB2500 Visual Chiseling".RosErrorNum := "DB2500 Visual Chiseling".RosErrorNum + 1; END_IF;
END_REGION

REGION Network 13: Step6: Read Page2 Point Data From ROS, then Save to DB | PLC Status Word:115 ROS Status Word: 215
   IF #High AND "DB2500 Visual Chiseling".VisualChiselingMode AND "DB2500 Visual Chiseling".VisualCameraStart AND ("DB2100 Modbus Value"."PLC Para"."Status Word" = 115) AND ("DB2100 Modbus Value"."ROS Para"."Status Word" = 215) AND ("DB2100 Modbus Value"."ROS Para"."PointPage Word" = 2) THEN
       #RetValue[10] := MOVE_BLK_VARIANT(SRC := P#DB2100.DBX0.0 BYTE 254,
                               COUNT := 144,
                               SRC_INDEX := 78,
                               DEST_INDEX := 0,
                               DEST => P#DB2300.DBX144.0 BYTE 288);
   END_IF;
END_REGION

REGION Network 14: Step6: Confirm Page2 Points Data Has been Received | PLC Status Word:120
   "Timer25_ChiselPage2".TON(IN := #High AND "DB2500 Visual Chiseling".VisualChiselingMode AND "DB2500 Visual Chiseling".VisualCameraStart AND ("DB2100 Modbus Value"."PLC Para"."Status Word" = 115) AND ("DB2100 Modbus Value"."ROS Para"."Status Word" = 215) AND ("DB2100 Modbus Value"."ROS Para"."PointPage Word" = 2),
                           PT := T#0.5s);
   IF "Timer25_ChiselPage2".Q THEN "DB2100 Modbus Value"."PLC Para"."Status Word" := 120; END_IF;
   "DB2500 Visual Chiseling".Page1_ConfirmInf := "Timer25_ChiselPage2".Q;
END_REGION

REGION Network 15: Step6: Calculate ROS Error When Receiving Page2 Point Data | PLC Status Word:115 ROS Status Word: 99
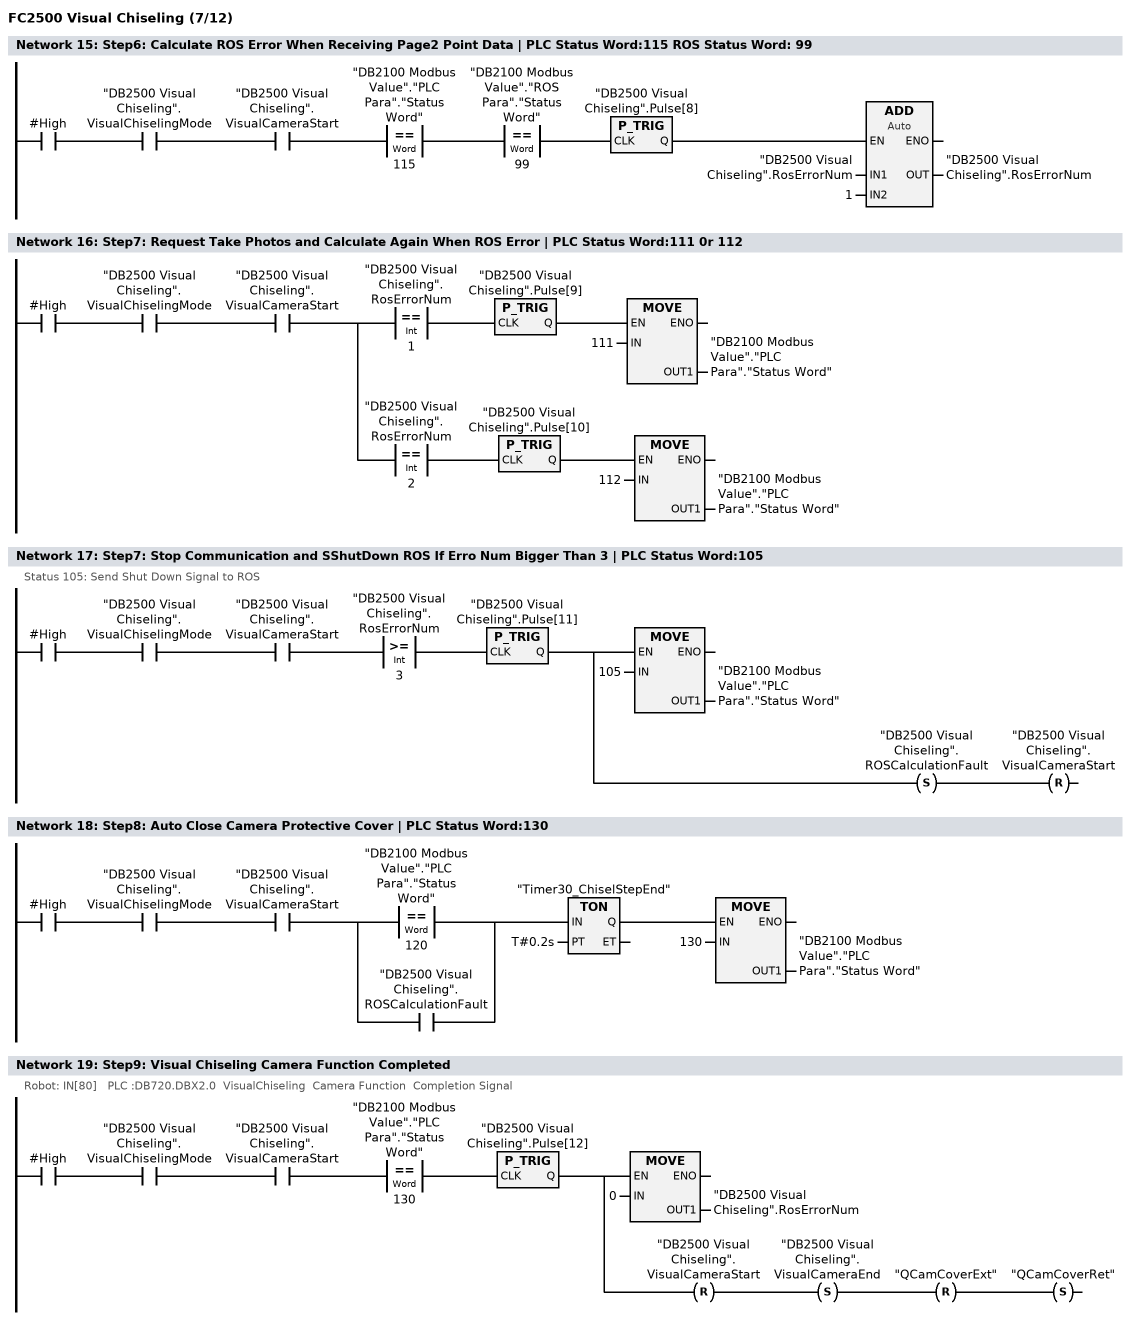
   RUNG wire#powerrail
      Contact( #High )
      Contact( "DB2500 Visual Chiseling".VisualChiselingMode )
      Contact( "DB2500 Visual Chiseling".VisualCameraStart )
      { S7_Templates := "SrcType := Word" } EQ_Contact(in1 := "DB2100 Modbus Value"."PLC Para"."Status Word", in2 := 115)
      { S7_Templates := "SrcType := Word" } EQ_Contact(in1 := "DB2100 Modbus Value"."ROS Para"."Status Word", in2 := 99)
      P_Trig( "DB2500 Visual Chiseling".Pulse[8] )
      Add(in1 := "DB2500 Visual Chiseling".RosErrorNum, in2 := 1, out => "DB2500 Visual Chiseling".RosErrorNum)
   END_RUNG
   // the same network as SCL:
   #_w1 := #High AND "DB2500 Visual Chiseling".VisualChiselingMode AND "DB2500 Visual Chiseling".VisualCameraStart AND ("DB2100 Modbus Value"."PLC Para"."Status Word" = 115) AND ("DB2100 Modbus Value"."ROS Para"."Status Word" = 99);
   #_w2 := #_w1 AND NOT "DB2500 Visual Chiseling".Pulse[8];   // rising edge
   "DB2500 Visual Chiseling".Pulse[8] := #_w1;
   IF #_w2 THEN "DB2500 Visual Chiseling".RosErrorNum := "DB2500 Visual Chiseling".RosErrorNum + 1; END_IF;
END_REGION

